(* IEC 61131-3 sources: JingjiangArm/moonboxpro_arm_8.4/Application/Application/任务列表/Main_Task/横向调整处理, 17 files *)

(* ---- StDigitalMicroStepDrive.st ---- *)
(*@CES
Name=StDigitalMicroStepDrive
Type=Gvl
TypeGuid=2db5746d-d284-4425-9f7f-2663a34b0ebc
Guid=10e217d5-ea4e-41f0-93bf-b76d90085cfe
HasDeclaration=True
HasImplementation=False
*)
{DECLARATION}
TYPE StDigitalMicroStepDrive :(*步进电机结构体*)
STRUCT
	xStepDriveEn:BOOL;(*步进电机使能*)
	xStepDriveDir:BOOL;(*步进电机方向*)
	xStepDriveMode:BOOL;(*电机速度位置模式*)(*TRUE 为位置模式，false为速度模式*)
	xStepDriveSpeedMode_Run:BOOL;(*步进电机速度模式启动标志*)
	xStepDriveWorking:BOOL;(*脉冲输出中*)
	xStepDriveAlarm:BOOL;(*步进电机报警*)
	iStepDriveState:INT;(*步进电机状态机*)

	udiStepDriveWorkingTime:UDINT;(*步进电机执行时间*)
	iStepDrivePulsePRev:INT;(*步进电机每圈的脉冲数*)
	iStepDriveNum:INT;(*步进电机减速比分子*)
	iStepDriveDen:INT;(*步进电机减速比分母*)
	lrStepDrivePosPPulse:LREAL;(*步进电机每个脉冲对应的位置值，单位mm*)(*通过测量得到，或者通过计算得到*)
	iStepDriveAccTime_ms:INT;(*步进电机加速时间ms*)
	wStepDrivePulseFre_Sa:WORD;(*步进电机启动脉冲频率*)
	wStepDrivePulseFre_Tar:WORD;(*步进电机目标脉冲频率*)
	wStepDriveAcc_SaToTar:WORD;(*到达目标速度的加速度*)
	wStepDrivePulse:WORD;(*步进电机脉冲数*)
	diStepDrivePluse_Act:DINT;(*步进电机实际走的脉冲数*)
	wStepDrivePulse_Act_Rd_Bak:WORD;(*读取到的步进电机上个周期实际走的脉冲数*)

(*读取模块中的数据*)
	awSpace:ARRAY [1..3] OF WORD;(*W0,W1,W2*)
	wStepDrivePulse_Act_Rd:WORD;(*读取到的步进电机实际走的脉冲数*)(*W3*)
	wStepDriveModuleIOData_Rd:WORD;(*步进电机模块的io输入值*)(*W4*)
	wStepDriveCTL_Rd:WORD;(*读取到的模块的数据*)(*W5*)
(*写入到模块中的参数。规定使用数字量模块 但是plc配置的时候需要配置模拟量模块*)
	wStepDrivePulseFre_Sa_Wr:WORD;(*步进电机启动脉冲频率写入值*)(*W0*)
	wStepDrivePulseFre_Tar_Wr:WORD;(*步进电机目标脉冲频率写入值*)(*W1*)
	wStepDriveAcc_SaToTar_Wr:WORD;(*到达目标速度的加速度写入值*)(*W2*)
	wStepDrivePulse_Wr:WORD;(*步进电机脉冲数写入值*)(*W3*)
	wStepDriveModuleIOData_Wr:WORD;(*步进电机模块的io输出写入*)(*W4*)
	wStepDriveCTL:WORD;(*步进电机控制位*)(*bit9:反馈脉冲数清零(*W5*)
								bit10:脉冲输出标志，1：输出中
								bit11:电机方向
								bit12:速度模式时，高电平输出脉冲，低电平停止输出
								bit13:位置模式时，上升沿开始输出脉冲，脉冲个数到达时停止输出
								bit14:速度、位置模式 0：速度模式，1：位置模式
								bit15:模块使能 0：脉冲输出无效，1：有效
							        *)
END_STRUCT
END_TYPE

{IMPLEMENTATION}

(* ---- StEnc0410R.st ---- *)
(*@CES
Name=StEnc0410R
Type=Gvl
TypeGuid=2db5746d-d284-4425-9f7f-2663a34b0ebc
Guid=6f80462c-d6b3-455f-883a-2142632bafb1
HasDeclaration=True
HasImplementation=False
*)
{DECLARATION}
TYPE StEnc0410R :
STRUCT
	wInputModeCfg:WORD;(*模块输入配置*)
	wInputEncValue:WORD;(*模块输入的编码器个数*)
	wInputEncValue_Bak:WORD;(*上个周期模块输入的编码器个数*)
	diInputEncValue_Total:DINT;(*总的编码器输入个数*)
	diEncValue_Middle:DINT;(*中位临时值*)

	byEnc0410RInPutMode:BYTE;(*模块输入方式选择 0:正交脉冲 1:脉冲+方向 2:正负脉冲*)
	xEnc0410RInPutPulDir:BOOL;(*模块输入脉冲方向 TRUE 取反*)
	byEnc0410RInPutPulCntWay:BYTE;(*模块输入脉冲计数方式 0:z信号开始 1:一直计数*)
	byEncO410RInputVol:BYTE;(*模块输入的电压类型*)

	byEnc0410ROutPutMode:BYTE;(*模块是输出方式选择0:正交脉冲 1:脉冲+方向 2:正负脉冲*)
END_STRUCT
END_TYPE

{IMPLEMENTATION}

(* ---- StStepDriveIOModule.st ---- *)
(*@CES
Name=StStepDriveIOModule
Type=Gvl
TypeGuid=2db5746d-d284-4425-9f7f-2663a34b0ebc
Guid=050a5971-e7ba-4c31-b40e-01a320b97a7e
HasDeclaration=True
HasImplementation=False
*)
{DECLARATION}
TYPE StStepDriveIOModule :
STRUCT
	wIX:WORD;(*输入数据*)(*0：15位为数字量输入*)
	wQX:WORD;(*输出数据*)(*2：9位为数字量继电器输出位*)
END_STRUCT
END_TYPE

{IMPLEMENTATION}

(* ---- TypeEnumEncModule.st ---- *)
(*@CES
Name=TypeEnumEncModule
Type=Gvl
TypeGuid=2db5746d-d284-4425-9f7f-2663a34b0ebc
Guid=5080d035-0ec5-4151-a1b0-b148bbf57879
HasDeclaration=True
HasImplementation=False
*)
{DECLARATION}
TYPE TypeEnumEncModule :
(
	(*0:继电器数字量模块HCB5-1610-DRA*)
	ENCMODULE_HCB5_1610_DRA:=0,
	(*1:Enc0410R模块输出*)
	ENCMODULE_ENC0410R:=1
);
END_TYPE

{IMPLEMENTATION}

(* ---- TypeEnumStepDriveStat.st ---- *)
(*@CES
Name=TypeEnumStepDriveStat
Type=Gvl
TypeGuid=2db5746d-d284-4425-9f7f-2663a34b0ebc
Guid=3c3a1540-5152-4e9f-b7fc-bae736162d3c
HasDeclaration=True
HasImplementation=False
*)
{DECLARATION}
TYPE TypeEnumStepDriveStat :
(
	STEPDRIVE_IDLE,(*空闲*)
	STEPDRIVE_RUN,(*启动*)
	STEPDRIVE_CLR,(*状态清除*)
	STEPDRIVE_WAITING,(*等待一个周期*)
	STEPDRIVE_MODULE_VALID,(*模块使能*)
	STEPDRIVE_PULSEOUT,(*脉冲输出*)
	STEPDRIVE_ALARM(*报警*)
);
END_TYPE

{IMPLEMENTATION}

(* ---- KS_GetEncPluse.st ---- *)
(*@CES
Name=KS_GetEncPluse
Type=FunctionBlock
TypeGuid=6f9dac99-8de1-4efc-8465-68ac443b7d08
Guid=2bf59e22-f994-4ac5-8b2b-a54b74aea4c6
HasDeclaration=True
HasImplementation=True
*)
{DECLARATION}
FUNCTION KS_GetEncPluse : BOOL
VAR_INPUT
	i_pastStDigitalMicroStepDrive :POINTER TO ARRAY [1..MAX_UNIT_NUM] OF StDigitalMicroStepDrive;
	i_pastStEnc0410R:POINTER TO ARRAY [1..MAX_UNIT_NUM] OF StEnc0410R;
END_VAR
VAR
	iN: INT;
END_VAR

{IMPLEMENTATION}
IF i_pastStDigitalMicroStepDrive<>0 AND i_pastStEnc0410R<>0 THEN
	FOR iN:=1 TO MAX_UNIT_NUM BY 1 DO(*针对所有轴进行读取*)
		i_pastStEnc0410R^[iN].wInputEncValue:=
		i_pastStDigitalMicroStepDrive^[iN].wStepDriveModuleIOData_Rd;(*读取回来的编码器脉冲个数，和数字量模块输入公用地址*)

		KS_GetPulse_Act(ADR(i_pastStEnc0410R^[iN].wInputEncValue),
						ADR(i_pastStEnc0410R^[iN].wInputEncValue_Bak),
						ADR(i_pastStEnc0410R^[iN].diInputEncValue_Total) );
	END_FOR
END_IF

(* ---- KS_GetHorizonManuAdj.st ---- *)
(*@CES
Name=KS_GetHorizonManuAdj
Type=FunctionBlock
TypeGuid=6f9dac99-8de1-4efc-8465-68ac443b7d08
Guid=d3a21ffb-1d17-434b-a6db-735f209d6991
HasDeclaration=True
HasImplementation=True
*)
{DECLARATION}
FUNCTION KS_GetHorizonManuAdj : INT(*界面手动调整量2018.9.4.093836*)(*um*)(*返回值为实际需要调整的量，-22222为参数异常*)
(*2022.2.18.164444 按钮方向方向和运动方向相关了*)
(*增加了注释文字@正值是向操作侧@负值是向传动侧@已经和电机旋转方向相关了*)
(*2023.3.9.225628 通过查看动态库发现,动态库中将原来的左按钮赋值为otostudio约定的右按钮
右按钮赋值为otostudio的左按钮
@以前约定向左pabyHorManuBtn= 1 2 5
@向右pabyHorManuBtn=3 4 6
为了不修改动态库,在这里再进行一次取反以保证一致！！@将i_xHorManuDirSwitch=true*)
(*2024.11.6.093600 同步*)
(*2024.11.5.110659*)
(*重新处理界面手动按钮清理，防止整体清除界面手动按钮时B系被A系清理掉了*)
VAR_INPUT
	i_xHorManuDirSwitch:BOOL;(*方向取反*)
	i_iHorManuAdj_Step:INT;(*横向手动调整当量um*)
	i_iHorManuAdj_FastStep:INT;(*横向手动快速调整当量um*)
	i_iHorManuAdj_MidStep:INT;(*横向手动快速调整当量um*)
	piUnitId:POINTER TO INT;(*色组号*)

	pabyHorManuBtn:POINTER TO ARRAY [1..MAX_UNIT_NUM] OF BYTE;(*横向手动按钮，0为不调整，1为左向慢调0.05mm，2为左向快调暂定为0.5mm；3为右向慢调，4为右向快调；
										这里界面上的按钮只控制左右，逻辑控制横向电机是向传动侧还是操作侧运动*)
	padiHorAdjustMent:POINTER TO ARRAY [1..MAX_UNIT_NUM] OF DINT;(*横向手动调整的量*)
	i_iGrpAxisNum_Pu:INT;
	i_abyGrpAxisList: ARRAY [1..MAX_UNIT_NUM] OF BYTE; (*系的轴列表*)
	i_pstStSysParam: POINTER TO StSysParam;
END_VAR
VAR
	iN: INT;
	iCoeff: INT;(*方向系数*)
	iResult: INT;
	iUnitId: INT;
END_VAR

{IMPLEMENTATION}
KS_GetHorizonManuAdj:=0;
IF pabyHorManuBtn<>0 AND padiHorAdjustMent<>0 AND piUnitId<>0 THEN(*指针合法性检查*);
ELSE
	KS_GetHorizonManuAdj:=-22222;(*特殊值标识报警*)
	RETURN;
END_IF

piUnitId^:=0;
IF i_iHorManuAdj_Step<=0 THEN
	i_iHorManuAdj_Step:=50;(*0.05MM*)
ELSE;
END_IF

IF i_iHorManuAdj_FastStep<=0 THEN
	i_iHorManuAdj_FastStep:=500;(*0.5MM*)
ELSE;
END_IF
(*2022.8.9.094516处理0.02档位*)
IF i_iHorManuAdj_MidStep<=0 THEN
	i_iHorManuAdj_FastStep:=100;(*0.1MM*)
ELSE;
END_IF
(*一个周期只处理一个轴*)(*调整量的正值代表向操作侧运动*)
(*2021.10.26.091200  使用轴列表变量*)
FOR iUnitId:=1 TO i_iGrpAxisNum_Pu BY 1 DO(*检查所有色组*)
	iN:=i_abyGrpAxisList[iUnitId];
(*方向*)
	iCoeff:=0;
(*增加0.02档位2022.8.9.094247||*)
(*	IF  pabyHorManuBtn^[iN]=1 OR  pabyHorManuBtn^[iN]=2  THEN(*向左*)*)
	IF  pabyHorManuBtn^[iN]=1 OR  pabyHorManuBtn^[iN]=2 OR  pabyHorManuBtn^[iN]=5 THEN(*向左*)
		IF i_pstStSysParam^.astStUnitParam_UnSave[iN].xMotRev_PrnRoller THEN (*电机反转*)(*向左是向传动侧运动*)
			iCoeff:=-1;
		ELSE(*电机正转*)(*向左是向操作侧运动*)
			iCoeff:=1;
		END_IF
	ELSIF  pabyHorManuBtn^[iN]=3 OR  pabyHorManuBtn^[iN]=4 OR  pabyHorManuBtn^[iN]=6 THEN (*向右*)(*和向左取反*)
		IF i_pstStSysParam^.astStUnitParam_UnSave[iN].xMotRev_PrnRoller THEN (*电机反转*)
			iCoeff:=1;
		ELSE(*电机正转*)
			iCoeff:=-1;
		END_IF
	END_IF

	IF i_xHorManuDirSwitch THEN
		iCoeff:=-iCoeff;
	END_IF
(*调整量值*)
	iResult:=0;
	IF  pabyHorManuBtn^[iN]=1 OR  pabyHorManuBtn^[iN]=3 THEN (*都是慢调*)
		iResult:=(i_iHorManuAdj_Step);
	ELSIF pabyHorManuBtn^[iN]=2 OR  pabyHorManuBtn^[iN]=4 THEN (*都是快调*)
		iResult:=(i_iHorManuAdj_FastStep);
	ELSIF pabyHorManuBtn^[iN]=5 OR  pabyHorManuBtn^[iN]=6 THEN (*中间档位-202022.8.9.094640*)
		iResult:=(i_iHorManuAdj_MidStep);
	END_IF
	iResult:=iResult*iCoeff;

	IF i_pstStSysParam^.astStUnitParam_Save[iN].xLinkage THEN (*检查联动轴*)
		IF pabyHorManuBtn^[iN]<>0 THEN (*说明有调整按下了*)
			pabyHorManuBtn^[iN]:=0;(*清零按钮标志*)(*2024.11.5.110459*)
			KS_GetHorizonManuAdj:=iResult;(*将调整量输出*)
			piUnitId^:=iN;
			padiHorAdjustMent^[iN]:=padiHorAdjustMent^[iN]+iResult;(*在界面显示*)
			EXIT;
		END_IF
	ELSE
		pabyHorManuBtn^[iN]:=0;(*清零按钮标志*)(*2024.11.5.110459*)
	END_IF
END_FOR

(* ---- KS_GetPulse_Act.st ---- *)
(*@CES
Name=KS_GetPulse_Act
Type=FunctionBlock
TypeGuid=6f9dac99-8de1-4efc-8465-68ac443b7d08
Guid=7e51e991-78cc-4457-be42-c8156f7134b7
HasDeclaration=True
HasImplementation=True
*)
{DECLARATION}
FUNCTION KS_GetPulse_Act : int
VAR_INPUT
	pwStepDrivePulse_Act_Rd :POINTER TO WORD;(*读取到的脉冲数*)
	pwStepDrivePulse_Act_Rd_Bak:POINTER TO WORD;(*上个周期读到的脉冲数*)
	pdiStepDrivePulse_Act:POINTER TO DINT;(*实际走的脉冲数*)
END_VAR
VAR
	iStepDrivePulse_Act_Rd: INT;
	iStepDrivePulse_Act_Rd_Bak: INT;
	iDeltaPulse: INT;(*步进电机脉冲变化量*)
END_VAR

{IMPLEMENTATION}
KS_GetPulse_Act:=0;
IF pwStepDrivePulse_Act_Rd<>0 AND pwStepDrivePulse_Act_Rd_Bak<>0 AND pdiStepDrivePulse_Act <>0 THEN;
ELSE
	KS_GetPulse_Act:=-1;
	RETURN;
END_IF

iStepDrivePulse_Act_Rd:=WORD_TO_INT(pwStepDrivePulse_Act_Rd^);
iStepDrivePulse_Act_Rd_Bak:= WORD_TO_INT(pwStepDrivePulse_Act_Rd_Bak^);

IF iStepDrivePulse_Act_Rd <> iStepDrivePulse_Act_Rd_Bak THEN
	iDeltaPulse:=(iStepDrivePulse_Act_Rd-iStepDrivePulse_Act_Rd_Bak);
	pdiStepDrivePulse_Act^:=pdiStepDrivePulse_Act^+iDeltaPulse;
ELSE;
END_IF

pwStepDrivePulse_Act_Rd_Bak^:=INT_TO_WORD(iStepDrivePulse_Act_Rd);(*保存上个周期的值*)

(* ---- KS_SetStepDriveModulePara.st ---- *)
(*@CES
Name=KS_SetStepDriveModulePara
Type=FunctionBlock
TypeGuid=6f9dac99-8de1-4efc-8465-68ac443b7d08
Guid=21a3679d-2e4f-4802-b9d7-d00f676e215d
HasDeclaration=True
HasImplementation=True
*)
{DECLARATION}
FUNCTION KS_SetStepDriveModulePara : BOOL(*设置步进电机脉冲输出模块脉冲方式参数*)
(*2019.5.15.112350|liu.yt|必须放在KS_FB_StepDriveCTL后执行，KS_FB_StepDriveCTL会清零，功能块再次再次赋值，反之则无效赋值*)
(*2019.4.18.130455 增加了ENCO410R型模块输入输出控制参数,主要用于高速编码器输入输出控制。MHZ频率*)
VAR_INPUT
	i_xMultiple_Input: BOOL;(*参数输入方式选择：多参数 或者 单参数*)
	i_byEncO410RInputVol:BYTE;(*模块输入的电压类型选择：0 是5v；1是24v*)
	i_byEnc0410RInPutMode:BYTE;(*模块输入方式选择 0:正交脉冲 1:脉冲+方向 2:正负脉冲*)
	i_xEnc0410RInPutPulDir:BOOL;(*模块输入脉冲方向 TRUE 取反*)
	i_byEnc0410RInPutPulCntWay:BYTE;(*模块输入脉冲计数方式 0:z信号开始 1:一直计数*)

	i_byEnc0410ROutPutMode:BYTE;(*模块输出方式选择 0:正交脉冲 1:脉冲+方向 2:正负脉冲*)
	i_pastStDigitalMicroStepDrive :POINTER TO ARRAY [1..MAX_UNIT_NUM] OF StDigitalMicroStepDrive;
	i_pastStEnc0410R:POINTER TO ARRAY [1..MAX_UNIT_NUM] OF StEnc0410R;
END_VAR
VAR
(*bit7:8 脉冲输出模式，仅限于EncO410R模块，0:正交脉冲 1:脉冲+方向 2:正负脉冲*)
	wEncO410ROutPutMode_ClrCtlBit:WORD:=16#FE7F;(*利用与运算清除7:8位*)
(*利用或运算定义控制位*)
	wEncO410ROutPutMode_QuadPul:WORD:=0;		(*正交脉冲输出模式	bit 7:8=0*)
	wEncO410ROutPutMode_PulAndDir:WORD:=16#0080;	(*脉冲+方向输出模式	bit 7:8=1*)
	wEncO410ROutPutMode_PlusMinusPul:WORD:=16#0100;(*正负脉冲输出模式	bit 7:8=2*)

(*************************************************)
(*Enc0410R 模块输入配置*)(*bit0:1 脉冲输入模式。bit2 方向取反。bit3 计数模式*)
	wEncO410RInPutMode_ClrCtlBit:WORD:=16#FFF0;(*利用与运算清除低四位*)
(*利用或运算定义控制位*)
	wEncO410RInPutMode_QuadPul:WORD:=0;		(*正交脉冲输出模式	bit 0:1=0*)
	wEncO410RInPutMode_PulAndDir:WORD:=16#0001;	(*脉冲+方向输出模式	bit 0:1=1*)
	wEncO410RInPutMode_PlusMinusPul:WORD:=16#0002;(*正负脉冲输出模式	bit 0:1=2*)
	wEncO410RInPutMode_PlusDir:WORD:=16#0004;(*bit2 脉冲方向*)
(*	wEncO410RInPutMode_PlusCntWay_Z:WORD:=0;(*脉冲计数模式：z信号开始*)*)
	wEncO410RInPutMode_PlusCntWay_All:WORD:=16#0008;(*脉冲计数模式：一直计数*)
	wEncO410RInPutMode_Vol:WORD:=16#0010;(*bit4 电压输入类型 0 是5v；1是24v*)

	iN: INT;
	wStepDriveCTL: WORD;
	wEncO410RInPutModeCfg: WORD;

	byEnc0410RInPutMode:BYTE;(*模块输入方式选择 0:正交脉冲 1:脉冲+方向 2:正负脉冲*)
	xEnc0410RInPutPulDir:BOOL;(*模块输入脉冲方向 TRUE 取反*)
	byEnc0410RInPutPulCntWay:BYTE;(*模块输入脉冲计数方式 0:z信号开始 1:一直计数*)
	byEncO410RInputVol: BYTE;(*模块输入的电压类型选择：0 是5v；1是24v*)

	byEnc0410ROutPutMode:BYTE;(*模块输出方式选择 0:正交脉冲 1:脉冲+方向 2:正负脉冲*)
END_VAR

{IMPLEMENTATION}
IF i_pastStDigitalMicroStepDrive<>0 AND i_pastStEnc0410R<>0 THEN
	FOR iN:=1 TO MAX_UNIT_NUM BY 1 DO(*针对所有轴进行控制*)
		IF i_xMultiple_Input THEN(*多参数输入*)
			byEnc0410RInPutMode:=i_pastStEnc0410R^[iN].byEnc0410RInPutMode;
			xEnc0410RInPutPulDir:=i_pastStEnc0410R^[iN].xEnc0410RInPutPulDir;
			byEnc0410RInPutPulCntWay:=i_pastStEnc0410R^[iN].byEnc0410RInPutPulCntWay;
			byEncO410RInputVol:=i_pastStEnc0410R^[iN].byEncO410RInputVol;
			byEnc0410ROutPutMode:=i_pastStEnc0410R^[iN].byEnc0410ROutPutMode;
		ELSE(*单参数输入*)
			byEnc0410RInPutMode:=i_byEnc0410RInPutMode;
			xEnc0410RInPutPulDir:=i_xEnc0410RInPutPulDir;
			byEnc0410RInPutPulCntWay:=i_byEnc0410RInPutPulCntWay;
			byEncO410RInputVol:=i_byEncO410RInputVol;
			byEnc0410ROutPutMode:=i_byEnc0410ROutPutMode;
		END_IF

		(*脉冲输出配置*)
		wStepDriveCTL:=i_pastStDigitalMicroStepDrive^[iN].wStepDriveCTL;
		wStepDriveCTL:=wStepDriveCTL AND wEncO410ROutPutMode_ClrCtlBit;(*清零相应位*)
		(*输出方式配置*)
		CASE byEnc0410ROutPutMode OF
		1:(*脉冲+方向*)
			wStepDriveCTL:=wStepDriveCTL+wEncO410ROutPutMode_PulAndDir;
		2:(*正负脉冲*)
			wStepDriveCTL:=wStepDriveCTL+wEncO410ROutPutMode_PlusMinusPul;
		ELSE(*默认输出方式是正交脉冲*)
			wStepDriveCTL:=wStepDriveCTL+wEncO410ROutPutMode_QuadPul;
		END_CASE

		i_pastStDigitalMicroStepDrive^[iN].wStepDriveCTL:=wStepDriveCTL;

		(*脉冲输入配置*)
		(*Enc0410R的输入参数配置和继电器数字量模块公用IO输入输出地址*)
		wEncO410RInPutModeCfg:=0;

		(*输入方式配置*)

		CASE byEnc0410RInPutMode OF
		1:(*脉冲+方向*)
			wEncO410RInPutModeCfg:=wEncO410RInPutModeCfg+wEncO410RInPutMode_PulAndDir;
		2:(*正负脉冲*)
			wEncO410RInPutModeCfg:=wEncO410RInPutModeCfg+wEncO410RInPutMode_PlusMinusPul;
		ELSE(*默认输出方式是正交脉冲*)
			wEncO410RInPutModeCfg:=wEncO410RInPutModeCfg+wEncO410RInPutMode_QuadPul;
		END_CASE

		(*方向取反*)
		IF xEnc0410RInPutPulDir THEN wEncO410RInPutModeCfg:=wEncO410RInPutModeCfg+wEncO410RInPutMode_PlusDir;END_IF

		(*计数方式选择*)
		IF byEnc0410RInPutPulCntWay<>0 THEN wEncO410RInPutModeCfg:=wEncO410RInPutModeCfg+wEncO410RInPutMode_PlusCntWay_All;END_IF

		(*输入电压类型 0 是5v  1是24v*)
		IF byEncO410RInputVol=1 THEN wEncO410RInPutModeCfg:=wEncO410RInPutModeCfg+wEncO410RInPutMode_Vol;END_IF

		i_pastStEnc0410R^[iN].wInputModeCfg:=wEncO410RInPutModeCfg;
	END_FOR
END_IF

(* ---- KS_FB_AxisHorAdj.st ---- *)
(*@CES
Name=KS_FB_AxisHorAdj
Type=FunctionBlock
TypeGuid=6f9dac99-8de1-4efc-8465-68ac443b7d08
Guid=bd4bc8d3-26df-4dfe-bfb9-1ac44a7e80cd
HasDeclaration=True
HasImplementation=True
*)
{DECLARATION}
FUNCTION_BLOCK KS_FB_AxisHorAdj(*从站横向*)
(*2022.6.10.161033 修复横向运动限位问题*)
(*屏蔽使用移动到KS_FB_GrpHorAdj函数中*)
(*2025.4.20.104124从站横向运动功能，停机状态取消联动相关|开机状态下非联动轴也可以运动*)
(*已经不使用了@@@@*)
VAR_INPUT
	i_xEn									: BOOL;(*功能块使能*)
	i_iGrpAxisNum_Pu						: INT; (*色组轴数*)
	i_aiGrpAxisList							: ARRAY [1..MAX_UNIT_NUM] OF INT; (*系的轴列表*)
	i_pastStIOMap_AxisBasic					: POINTER TO ARRAY [1..MAX_UNIT_NUM] OF StIOMap_Axis_FE; (*基础io|*)
	i_xFlag_Estop							: BOOL;(*急停标志*)
	i_xFlag_Stop							: BOOL;(*停机标志*)
	i_lrVel_HorzPreRegister					: LREAL;
	i_lrVel_HorzAdjust						: LREAL;
	i_iCycleTime_Plc						: INT;
	i_pastStAxisRapidAdjProf_H				: POINTER TO ARRAY [1..MAX_UNIT_NUM] OF StAxisRapidAdjProf_H;(*纵向快速对版|*)
	i_pstStSysParam: POINTER TO StSysParam;
	i_iGrpId: INT;
END_VAR
VAR_OUTPUT

	o_axAxisHorAdjing: ARRAY [1..MAX_UNIT_NUM] OF BOOL;
END_VAR
VAR
	iN: INT;
	iUnitId: INT;
	//pstStAxisParam: POINTER TO StAxisParam;
	pstStIOMap_AxisBasic: POINTER TO StIOMap_Axis_FE;

	lrAdjustVal_H_PerCycle: LREAL;
	axAxisHorAdjSts: ARRAY [1..MAX_UNIT_NUM] OF BOOL;
	axAxisHorAdj_End: ARRAY [1..MAX_UNIT_NUM] OF BOOL;
	iRtn: INT;
	iAdjustment_HorAxisAdj: INT;
	axHorAxisAdjStop: ARRAY [1..MAX_UNIT_NUM] OF BOOL;
	axHorAxisAdjStart: ARRAY [1..MAX_UNIT_NUM] OF BOOL;
	xFlag_HorAxisAdj: BOOL;
	wSts_HorzManuPreReg:WORD;
	xAutoMove_H: BOOL;(*2025.4.20.110020+*)
END_VAR

{IMPLEMENTATION}
IF i_xEn AND
	(i_iGrpAxisNum_Pu>=1 AND i_iGrpAxisNum_Pu<=MAX_UNIT_NUM) AND
	i_pastStIOMap_AxisBasic<>0 AND
	i_pastStAxisRapidAdjProf_H<>0 THEN(*2019.11.18.153726_*)

	FOR iN:= 1 TO i_iGrpAxisNum_Pu BY 1 DO
		iUnitId:= i_aiGrpAxisList[iN];
		pstStIOMap_AxisBasic:= ADR(i_pastStIOMap_AxisBasic^[iUnitId]);

		(*--------------------------------------------------|2019.11.18.153930_*)
		(*横向快速对版改成单个轴处理时放在循环内处理|*)
		iRtn:= KS_FetchRapidAdjValue_H(i_pastStAxisRapidAdjProf_H, iUnitId, ADR(iAdjustment_HorAxisAdj));
		(*2025.4.20.110359 同步*)
		(*2024.01.17.161205 增加清除处理*)
		axHorAxisAdjStart[iUnitId]:= FALSE;
		axHorAxisAdjStop[iUnitId]:= FALSE;
		IF iRtn=0 THEN
			IF iAdjustment_HorAxisAdj=-32767 THEN(*人为停止标志|*)
				axHorAxisAdjStop[iUnitId]:= TRUE;
				axHorAxisAdjStart[iUnitId]:= FALSE;
			ELSIF iAdjustment_HorAxisAdj<>0 THEN
				axHorAxisAdjStop[iUnitId]:= FALSE;
				axHorAxisAdjStart[iUnitId]:= TRUE;
				i_pstStSysParam^.astStUnitParam_UnSave[iUnitId].alrTotalAdjustVal_ManuCoarse_vh[2]:= i_pstStSysParam^.astStUnitParam_UnSave[iUnitId].alrTotalAdjustVal_ManuCoarse_vh[2]+iAdjustment_HorAxisAdj;
			END_IF
		END_IF

		IF (NOT i_xFlag_Estop) (*AND i_xFlag_Stop*) THEN(*非急停*)
			(*2025.4.20.105720 修改条件*)
			IF i_xFlag_Stop THEN(*不用限制单联动*)
				xAutoMove_H:=TRUE;
			ELSE(*非停机状态下|只有单动的可以*)
				xAutoMove_H:=NOT i_pstStSysParam^.astStUnitParam_Save[iUnitId].xLinkage;
			END_IF

			IF (*pstStAxisParam^.xLinkage*)xAutoMove_H THEN
				IF axHorAxisAdjStart[iUnitId] AND (NOT axAxisHorAdjSts[iUnitId]) THEN(*开始运行*)
					axAxisHorAdjSts[iUnitId]:= TRUE;
					axHorAxisAdjStart[iUnitId]:= FALSE;
				END_IF
				IF axHorAxisAdjStop[iUnitId] AND axAxisHorAdjSts[iUnitId] THEN(*停止运行*)
					axAxisHorAdjSts[iUnitId]:= FALSE;
					axHorAxisAdjStop[iUnitId]:= FALSE;
				END_IF
			ELSE
				axHorAxisAdjStart[iUnitId]:= FALSE;
				axHorAxisAdjStop[iUnitId]:= FALSE;
				axAxisHorAdjSts[iUnitId]:= FALSE;
				IF i_pstStSysParam^.astStUnitParam_UnSave[iUnitId].alrTotalAdjustVal_ManuCoarse_vh[2]<>0 THEN
					i_pstStSysParam^.astStUnitParam_UnSave[iUnitId].alrTotalAdjustVal_ManuCoarse_vh[2]:= 0;
				END_IF

			END_IF
		ELSE(*2019.11.20.115512 增加了清除axHorAxisAdjStart
								axHorAxisAdjStop标志|Liu.yt*)
			axHorAxisAdjStart[iUnitId]:= FALSE;
			axHorAxisAdjStop[iUnitId]:= FALSE;
			IF axAxisHorAdjSts[iUnitId] THEN
				axAxisHorAdjSts[iUnitId]:= FALSE;(*急停或者非停机-直接停止运行*)
				i_pstStSysParam^.astStUnitParam_UnSave[iUnitId].alrTotalAdjustVal_ManuCoarse_vh[2]:= 0;
			END_IF
		END_IF

		IF pstStIOMap_AxisBasic^.o_xRel_Press OR (NOT pstStIOMap_AxisBasic^.i_xHorzMotor_FastSpd) THEN
		(*快调/慢调处理*)
			lrAdjustVal_H_PerCycle:= i_lrVel_HorzAdjust*INT_TO_LREAL(i_iCycleTime_Plc);
		ELSE
			lrAdjustVal_H_PerCycle:= i_lrVel_HorzPreRegister*INT_TO_LREAL(i_iCycleTime_Plc);
		END_IF

		IF axAxisHorAdjSts[iUnitId] THEN (*色组进入到横向对版状态*)
			xFlag_HorAxisAdj:= TRUE;

			(*2025.4.20.105821 屏蔽联动条件*)
			IF i_pstStSysParam^.astStUnitParam_Save[iUnitId].xLinkage OR TRUE THEN(*色组联动*)
				IF NOT axAxisHorAdj_End[iUnitId] THEN
					IF NOT o_axAxisHorAdjing[iUnitId] THEN
						o_axAxisHorAdjing[iUnitId]:= TRUE;
						(*横向对版量叠加到横向手动粗调仓库*)
						i_pstStSysParam^.astStUnitParam_UnSave[iUnitId].alrTotalAdjustVal_ManuCoarse_vh[2]:= -i_pstStSysParam^.astStUnitParam_UnSave[iUnitId].alrTotalAdjustVal_ManuCoarse_vh[2]*1000;(*单位um*)
					ELSE
(*2022.6.10.160946*)
(*
						IF pstStIOMap_AxisBasic^.i_xPosLimit_Left OR pstStIOMap_AxisBasic^.i_xPosLimit_Right THEN (*到达左右限位，直接清零调整量*)
							pstStAxisParam^.alrTotalAdjustVal_ManuCoarse_vh[2]:= 0;
						END_IF
*)

						IF (pstStIOMap_AxisBasic^.i_xPosLimit_Right AND i_pstStSysParam^.astStUnitParam_UnSave[iUnitId].alrTotalAdjustVal_ManuCoarse_vh[2]<0) OR
							(pstStIOMap_AxisBasic^.i_xPosLimit_Left AND i_pstStSysParam^.astStUnitParam_UnSave[iUnitId].alrTotalAdjustVal_ManuCoarse_vh[2]>0) THEN
							i_pstStSysParam^.astStUnitParam_UnSave[iUnitId].alrTotalAdjustVal_ManuCoarse_vh[2]:=0;
						END_IF

						IF i_pstStSysParam^.astStUnitParam_UnSave[iUnitId].alrTotalAdjustVal_ManuCoarse_vh[2]=0 THEN(*调整量消耗完成*)
							o_axAxisHorAdjing[iUnitId]:= FALSE;
							axAxisHorAdj_End[iUnitId]:= TRUE;
							axAxisHorAdjSts[iUnitId]:= FALSE;
						END_IF
					END_IF
				END_IF
			ELSE(*单动*)
				o_axAxisHorAdjing[iUnitId]:= FALSE;
				axAxisHorAdj_End[iUnitId]:= TRUE;
				axAxisHorAdjSts[iUnitId]:= FALSE;
				IF i_pstStSysParam^.astStUnitParam_UnSave[iUnitId].alrTotalAdjustVal_ManuCoarse_vh[2]<>0 THEN
					i_pstStSysParam^.astStUnitParam_UnSave[iUnitId].alrTotalAdjustVal_ManuCoarse_vh[2]:=0;
				END_IF
			END_IF
		ELSE
			IF xFlag_HorAxisAdj THEN
				xFlag_HorAxisAdj:= FALSE;
			END_IF
			o_axAxisHorAdjing[iUnitId]:= FALSE;
			axAxisHorAdj_End[iUnitId]:= FALSE;
			IF i_pstStSysParam^.astStUnitParam_UnSave[iUnitId].alrTotalAdjustVal_ManuCoarse_vh[2]<>0 THEN(*退出横向对版状态，调整量清零*)
				i_pstStSysParam^.astStUnitParam_UnSave[iUnitId].alrTotalAdjustVal_ManuCoarse_vh[2]:=0;
			END_IF
		END_IF

		IF axAxisHorAdjSts[iUnitId] THEN
			IF ABS(i_pstStSysParam^.astStUnitParam_UnSave[iUnitId].alrTotalAdjustVal_ManuCoarse_vh[2])>lrAdjustVal_H_PerCycle THEN
				IF i_pstStSysParam^.astStUnitParam_UnSave[iUnitId].alrTotalAdjustVal_ManuCoarse_vh[2]>0 THEN
					(*正向*)
					i_pstStSysParam^.astStUnitParam_UnSave[iUnitId].alrCurCycleAdjustVal_ManuCoarse_vh[2]:= lrAdjustVal_H_PerCycle;
					i_pstStSysParam^.astStUnitParam_UnSave[iUnitId].alrTotalAdjustVal_ManuCoarse_vh[2]:= i_pstStSysParam^.astStUnitParam_UnSave[iUnitId].alrTotalAdjustVal_ManuCoarse_vh[2] - i_pstStSysParam^.astStUnitParam_UnSave[iUnitId].alrCurCycleAdjustVal_ManuCoarse_vh[2];
					i_pstStSysParam^.astStUnitParam_UnSave[iUnitId].axCurCycleAdjustVal_ManuCoarse_done_vh[2]:= FALSE;
					pstStIOMap_AxisBasic^.o_xHorzMotor_CW:= TRUE;(*正转*)
					pstStIOMap_AxisBasic^.o_xHorzMotor_CCW:= FALSE;
				ELSE
					(*反向*)
					i_pstStSysParam^.astStUnitParam_UnSave[iUnitId].alrCurCycleAdjustVal_ManuCoarse_vh[2]:= -lrAdjustVal_H_PerCycle;
					i_pstStSysParam^.astStUnitParam_UnSave[iUnitId].alrTotalAdjustVal_ManuCoarse_vh[2]:= i_pstStSysParam^.astStUnitParam_UnSave[iUnitId].alrTotalAdjustVal_ManuCoarse_vh[2] - i_pstStSysParam^.astStUnitParam_UnSave[iUnitId].alrCurCycleAdjustVal_ManuCoarse_vh[2];
					i_pstStSysParam^.astStUnitParam_UnSave[iUnitId].axCurCycleAdjustVal_ManuCoarse_done_vh[2]:= FALSE;
					pstStIOMap_AxisBasic^.o_xHorzMotor_CCW:= TRUE;(*反转*)
					pstStIOMap_AxisBasic^.o_xHorzMotor_CW:= FALSE;
				END_IF
			ELSE
				IF o_axAxisHorAdjing[iUnitId] THEN
					i_pstStSysParam^.astStUnitParam_UnSave[iUnitId].alrTotalAdjustVal_ManuCoarse_vh[2]:= 0;
				END_IF
				pstStIOMap_AxisBasic^.o_xHorzMotor_CW:= FALSE;
				pstStIOMap_AxisBasic^.o_xHorzMotor_CCW:= FALSE;
			END_IF

		END_IF
(*往从站发送*)
		i_pstStSysParam^.astStUnitParam_UnSave[iUnitId].iPos_HorzManuPreReg:= -LREAL_TO_INT(i_pstStSysParam^.astStUnitParam_UnSave[iUnitId].alrTotalAdjustVal_ManuCoarse_vh[2]/1000);

		wSts_HorzManuPreReg.0:= o_axAxisHorAdjing[iUnitId];
		wSts_HorzManuPreReg.1:= pstStIOMap_AxisBasic^.o_xHorzMotor_CW;
		wSts_HorzManuPreReg.2:= pstStIOMap_AxisBasic^.o_xHorzMotor_CCW;
		wSts_HorzManuPreReg.3:= pstStIOMap_AxisBasic^.i_xPosLimit_Left;
		wSts_HorzManuPreReg.4:= pstStIOMap_AxisBasic^.i_xPosLimit_Right;
		wSts_HorzManuPreReg.5:= i_pstStSysParam^.astStGrpParam_UnSave[i_iGrpId].xFlag_Stop;

		i_pstStSysParam^.astStUnitParam_UnSave[iUnitId].wSts_HorzManuPreReg:= wSts_HorzManuPreReg;
	END_FOR

END_IF

(* ---- KS_FB_Debug_Get_mmPpul.st ---- *)
(*@CES
Name=KS_FB_Debug_Get_mmPpul
Type=FunctionBlock
TypeGuid=6f9dac99-8de1-4efc-8465-68ac443b7d08
Guid=61707722-1ee3-4896-b414-72dee3b67cb6
HasDeclaration=True
HasImplementation=True
*)
{DECLARATION}
FUNCTION_BLOCK KS_FB_Debug_Get_mmPpul(*调试模式下计算出的每个脉冲对应的位置值单位mm/pul*)
VAR_INPUT
	i_xEn:BOOL;(*功能块使能*)
	i_xStartTrig:BOOL;(*启动步进电机*)
	i_xCalEn:BOOL;(*计算使能标志*)
	i_iNum:INT;(*执行该动作的色组号*)
	i_iStepDriveSa_Vel:INT;(*步进电机启动速度*)
	i_iStepDrivePreReg_Vel:INT;(*z步进电机预套速度R/MIN*)
	i_diPulse:DINT;(*执行的脉冲数pul*)
	i_lrPos_Act:LREAL;(*实际走的距离mm*)
	i_pastStDigitalMicroStepDrive :POINTER TO ARRAY [1..MAX_UNIT_NUM] OF StDigitalMicroStepDrive;
END_VAR
VAR_OUTPUT
	o_xEn:BOOL;(**)
	o_xDebugTestDone: BOOL;(*测试完成了*)
	o_lrResult:LREAL;(*计算出的结果*)(*只有效一个周期*)
	o_iErrCode: INT;(*-1 地址错误。-2 数组下标越界,-3 输入参数错误*)
END_VAR
VAR
	xPreStartTrig: BOOL;(*用来控制启动检测按钮的上升沿*)
	stStDigitalMicroStepDrive_Temp: StDigitalMicroStepDrive;
	lrTemp: LREAL;
	lrTemp1: LREAL;
	xDebugTesting: BOOL;(*处于测试状态中*)
	xPreStepDriveWorking: BOOL;(*用来检测脉冲输出下降沿*)
	xPreCalEn: BOOL;(*用于检测计算使能上升沿*)
END_VAR

{IMPLEMENTATION}
(*输入参数检查*)
o_iErrCode:=0;
o_lrResult:=0;
IF i_pastStDigitalMicroStepDrive<>0 THEN;
ELSE
	o_iErrCode:=-1;
	RETURN;
END_IF

IF i_iNum>=1 AND i_iNum<=MAX_UNIT_NUM THEN
;
ELSE
	i_iNum:=1;
	o_iErrCode:=-2;
END_IF

IF ABS(i_diPulse)>65535 AND i_diPulse<>0 THEN
	i_diPulse:=65535*i_diPulse/i_diPulse;
	o_iErrCode:=-3;
END_IF

IF i_lrPos_Act<0 THEN
	i_lrPos_Act:=ABS(i_lrPos_Act);
	o_iErrCode:=-3;
END_IF

IF i_iStepDriveSa_Vel<0 THEN
	i_iStepDriveSa_Vel:=ABS(i_iStepDriveSa_Vel);
	o_iErrCode:=-3;
END_IF

IF i_iStepDrivePreReg_Vel<0 THEN
	i_iStepDrivePreReg_Vel:=ABS(i_iStepDrivePreReg_Vel);
	o_iErrCode:=-3;
END_IF

stStDigitalMicroStepDrive_Temp:=i_pastStDigitalMicroStepDrive^[i_iNum];
IF i_xEn THEN(*使能计算*)
	IF i_xStartTrig  AND NOT xPreStartTrig THEN(*检测按钮上升沿*)
		IF NOT xDebugTesting THEN
			o_xDebugTestDone:=FALSE;
			lrTemp:=i_pastStDigitalMicroStepDrive^[i_iNum].iStepDrivePulsePRev*i_iStepDriveSa_Vel/60.0;(*pul/s*)
			lrTemp1:=i_pastStDigitalMicroStepDrive^[i_iNum].iStepDrivePulsePRev*i_iStepDrivePreReg_Vel/60.0;(*pul/s*)
			IF i_pastStDigitalMicroStepDrive^[i_iNum].iStepDriveState=STEPDRIVE_IDLE  THEN(*空闲状态*)
				i_pastStDigitalMicroStepDrive^[i_iNum].iStepDriveState:=STEPDRIVE_RUN;(*启动步进电机调整*)
				i_pastStDigitalMicroStepDrive^[i_iNum].wStepDrivePulseFre_Sa:=LREAL_TO_WORD(lrTemp);
				i_pastStDigitalMicroStepDrive^[i_iNum].wStepDrivePulseFre_Tar:=LREAL_TO_WORD(lrTemp1);
				i_pastStDigitalMicroStepDrive^[i_iNum].wStepDrivePulse:=DINT_TO_WORD(ABS(i_diPulse));(*写入的脉冲数*)
				i_pastStDigitalMicroStepDrive^[i_iNum].xStepDriveMode:=TRUE;(*位置模式*)
				i_pastStDigitalMicroStepDrive^[i_iNum].xStepDriveSpeedMode_Run:=FALSE;(*置位速度模式输出标志*)
				IF i_diPulse>0 THEN
					i_pastStDigitalMicroStepDrive^[i_iNum].xStepDriveDir:=TRUE;(*为正值的时候我们认为是向传动侧转动，由于默认方向是向操作侧转动，故写为true*)
				ELSE
					i_pastStDigitalMicroStepDrive^[i_iNum].xStepDriveDir:=FALSE;(*为负值的时候我们认为是向操作侧转动，由于默认方向是向操作侧转动，故写为false*)
				END_IF
			END_IF
		ELSE(*再次按下启动按钮我们就退出测试位置的状态*);
			i_pastStDigitalMicroStepDrive^[i_iNum].iStepDriveState:=STEPDRIVE_IDLE;(*先退出到空闲状态*)
		END_IF
		xDebugTesting:=NOT xDebugTesting;
	END_IF

	IF xDebugTesting THEN (*已经处于测试的状态了,这个时候需要一直检测是否执行完成了*)
		IF NOT i_pastStDigitalMicroStepDrive^[i_iNum].xStepDriveWorking AND  xPreStepDriveWorking THEN(*脉冲输出标志下降沿*)
			i_pastStDigitalMicroStepDrive^[i_iNum].iStepDriveState:=STEPDRIVE_IDLE;(*退出到空闲状态*)
			xDebugTesting:=FALSE;
			o_xDebugTestDone:=TRUE;
		END_IF
	ELSE;
	END_IF

	IF o_xDebugTestDone THEN (*测试完成 接着我们计算每个脉冲对应的位置值*)
		IF i_xCalEn AND NOT xPreCalEn THEN(*计算上升沿标志*)
			IF i_pastStDigitalMicroStepDrive^[i_iNum].diStepDrivePluse_Act<>0 THEN
				o_lrResult:=ABS(i_lrPos_Act/i_pastStDigitalMicroStepDrive^[i_iNum].diStepDrivePluse_Act);
			ELSE
				o_iErrCode:=-4;
			END_IF
		END_IF
	END_IF
ELSE
	xDebugTesting:=FALSE;
	o_xDebugTestDone:=FALSE;
END_IF
xPreStepDriveWorking:=i_pastStDigitalMicroStepDrive^[i_iNum].xStepDriveWorking;
xPreStartTrig:=i_xStartTrig;
xPreCalEn:=i_xCalEn;

(* ---- KS_FB_GrpHorAdj.st ---- *)
(*@CES
Name=KS_FB_GrpHorAdj
Type=FunctionBlock
TypeGuid=6f9dac99-8de1-4efc-8465-68ac443b7d08
Guid=d546f829-7451-435f-8672-15bc73f9dc0f
HasDeclaration=True
HasImplementation=True
*)
{DECLARATION}
FUNCTION_BLOCK KS_FB_GrpHorAdj(*传统横向电机调整*)
(*2023.3.8.214754
移植KS_FB_AxisHorAdj 代码
程序逻辑只有操作侧和传动侧的方向
@位置正值代表向操作侧运动
@位置负值代表向传动侧运动
电机输出只有正转和反转
@正转是向操作侧
@反转是向传动侧*)
(*2023.3.10.105606 为了兼容外部的硬件限位处理
这里将限位定义调整下
@i_xMove_Left 为正转限位即操作侧限位
@i_xMove_Right 为反转限位即传动侧限位
@支持密码切换将限位定义切换为左右限位@dwControlComplexBits.17|未处理密码切换部分*)

(*2024.01.17.162016 优化从站横向控制标志处理@现场偶尔出现从站横向操作无响应问题*)
(*2025.4.20.104124从站横向运动功能，停机状态取消联动相关|开机状态下非联动轴也可以运动*)
(*2025.9.5.104845 自动横向调整时单周期调整量超过1丝的量不会因为自动速度太快而不响应@现场会出现小误差一直不能回来(单个周期的调整量太大了)*)
VAR_INPUT
	i_xEn: BOOL;(*使能*)
	i_iGrpAxisNum_Pu: INT; (*色组轴数*)
	i_abyGrpAxisList: ARRAY [1..MAX_UNIT_NUM] OF BYTE; (*系的轴列表*)
	i_pastStIOMap_AxisBasic: POINTER TO ARRAY [1..MAX_UNIT_NUM] OF StIOMap_Axis_FE; (*基础io|*)
	i_pastStIOMap_AxisExtra: POINTER TO ARRAY [1..MAX_UNIT_NUM] OF StIOMap_Axis_Extra_FE; (* 扩展io|*)
	i_lrVel_HorzAdjust		: LREAL;(*mm/s; um/ms; 横向调整速度|*)
	i_lrVel_HorzPreRegister		: LREAL;(*mm/s;横向预套准速度|*)
	(*2023.3.8.114628*)
	i_xFlag_Estop							: BOOL;(*急停标志*)
	i_xFlag_Stop							: BOOL;(*停机标志*)
	i_iCycleTime_Plc						: INT;
	i_pastStAxisRapidAdjProf_H				: POINTER TO ARRAY [1..MAX_UNIT_NUM] OF StAxisRapidAdjProf_H;(*纵向快速对版|*)
	i_pstStSysParam: POINTER TO StSysParam;
	i_xHorLimit:BOOL;(*横向限位定义修改为左右|默认是纤维定义为正反方向*)
	i_iGrpId: INT;
	i_xHorManuCtrl:BOOL;(*界面横向手动修正功能*)
END_VAR
VAR_OUTPUT
	o_xEno: BOOL;
	o_iErNo: INT;(*0成功\-1参数失败|*)
	o_axAxisHorAdjing: ARRAY [1..MAX_UNIT_NUM] OF BOOL;
END_VAR
VAR
	iN: INT;

	iUnitId: INT;

	pstStIOMap_AxisBasic: POINTER TO StIOMap_Axis_FE;
	pstStIOMap_AxisExtra: POINTER TO StIOMap_Axis_Extra_FE;
	//pstStAxisParam: POINTER TO StAxisParam;

	xFlag_PreRegister_H: BOOL;(*用来表征是否进入过横向预套准状态*)

	wHorzMotorDir: WORD;(*.0 |正转方向
					.1|反转方向*)
	awPreHorzMotorDir: ARRAY [1..MAX_UNIT_NUM] OF WORD;
	axHorzMotorStart_Delay: ARRAY [1..MAX_UNIT_NUM] OF BOOL;(*横向启动延时标志*)
	axHorzMotorStart_DelayDne: ARRAY [1..MAX_UNIT_NUM] OF BOOL;(*横向启动延时完成*)
	auiHorzMotorStart_Count: ARRAY [1..MAX_UNIT_NUM] OF UINT;(*启动延时计时变量*)
	iHorzMotorStart_DelayTime_MS: INT:=0;(*启动的延时时间ms*)

	adwTotalTimes_CW_AxisHorzManu: ARRAY [1..MAX_UNIT_NUM] OF DWORD ;
	adwTotalTimes_CCW_AxisHorzManu: ARRAY [1..MAX_UNIT_NUM] OF DWORD ;
	lrAdjustVal_H_PerCycle:LREAL;(*每个周期调整的量*)

	(*2023.3.8.114227 将函数KS_FB_AxisHorAdj中的代码移植到此处*)
	axAxisHorAdjSts: ARRAY [1..MAX_UNIT_NUM] OF BOOL;
	axAxisHorAdj_End: ARRAY [1..MAX_UNIT_NUM] OF BOOL;
	iRtn: INT;
	iAdjustment_HorAxisAdj: INT;
	axHorAxisAdjStop: ARRAY [1..MAX_UNIT_NUM] OF BOOL;
	axHorAxisAdjStart: ARRAY [1..MAX_UNIT_NUM] OF BOOL;
	xFlag_HorAxisAdj: BOOL;
	wSts_HorzManuPreReg:WORD;
	(*横向运动相关变量都使用操作侧和传动侧变量重新赋值@2023.3.8.104853*)
	axHorMovingBtn_M: ARRAY [1..MAX_UNIT_NUM] OF BOOL;(*横向操作侧运动按钮*)
	axHorMovingBtn_G: ARRAY [1..MAX_UNIT_NUM] OF BOOL;(*横向传动侧运动按钮*)
	axHorMovingLimit_M: ARRAY [1..MAX_UNIT_NUM] OF BOOL;(*横向操作侧运动限位*)
	axHorMovingLimit_G: ARRAY [1..MAX_UNIT_NUM] OF BOOL;(*横向传动侧运动限位*)
	axHorMoving_M: ARRAY [1..MAX_UNIT_NUM] OF BOOL;(*横向操作侧运动*)
	axHorMoving_G: ARRAY [1..MAX_UNIT_NUM] OF BOOL;(*横向传动侧运动*)
	xAutoMove_H: BOOL;(*2025.4.20.110711+*)
END_VAR

{IMPLEMENTATION}
o_xEno:= i_xEn;
o_iErNo:= 0;
IF i_xEn THEN
	IF (i_iGrpAxisNum_Pu>=1 AND i_iGrpAxisNum_Pu<=MAX_UNIT_NUM) AND(*系的色组数量有效|*)
		i_pastStIOMap_AxisBasic<>0 AND
		i_pastStIOMap_AxisExtra<>0 THEN

		(*2023.3.8.114227 将函数KS_FB_AxisHorAdj中的代码移植到此处*)
		FOR iN:= 1 TO i_iGrpAxisNum_Pu BY 1 DO
			iUnitId:= i_abyGrpAxisList[iN];
			pstStIOMap_AxisBasic:= ADR(i_pastStIOMap_AxisBasic^[iUnitId]);

			(*处理横向开关相关@2023.3.8.104924*)
			(*和运动方向关联@伺服正转(正手机)-左对应操作侧#先不关心反印时候的方向变化问题
						    @伺服反转(反手机)-左对应传动侧#先不关心反印时候的方向变化问题*)
			IF NOT i_pstStSysParam^.astStUnitParam_UnSave[iUnitId].xMotRev_PrnRoller THEN(*正转*)
				axHorMovingBtn_M[iUnitId]:=pstStIOMap_AxisBasic^.i_xMove_Left;
				axHorMovingBtn_G[iUnitId]:=pstStIOMap_AxisBasic^.i_xMove_Right;

				axHorMovingLimit_M[iUnitId]:=pstStIOMap_AxisBasic^.i_xPosLimit_Left;
				axHorMovingLimit_G[iUnitId]:=pstStIOMap_AxisBasic^.i_xPosLimit_Right;
			ELSE(*反转*)
				axHorMovingBtn_M[iUnitId]:=pstStIOMap_AxisBasic^.i_xMove_Right;
				axHorMovingBtn_G[iUnitId]:=pstStIOMap_AxisBasic^.i_xMove_Left;

				IF i_xHorLimit THEN
					(*使用左右限位*)
					axHorMovingLimit_M[iUnitId]:=pstStIOMap_AxisBasic^.i_xPosLimit_Right;
					axHorMovingLimit_G[iUnitId]:=pstStIOMap_AxisBasic^.i_xPosLimit_Left;
				ELSE
					(*使用正转(操作侧)反转(传动侧)限位*)
					axHorMovingLimit_M[iUnitId]:=pstStIOMap_AxisBasic^.i_xPosLimit_Left;
					axHorMovingLimit_G[iUnitId]:=pstStIOMap_AxisBasic^.i_xPosLimit_Right;
				END_IF
			END_IF

			(*--------------------------------------------------|2019.11.18.153930_*)
			(*横向快速对版改成单个轴处理时放在循环内处理|*)
			(*返回的距离单位是mm*)
			iAdjustment_HorAxisAdj:=0;(*清零*)
			iRtn:= KS_FetchRapidAdjValue_H(i_pastStAxisRapidAdjProf_H, iUnitId, ADR(iAdjustment_HorAxisAdj));
			(*2024.01.17.161205 增加清除处理*)
			axHorAxisAdjStart[iUnitId]:= FALSE;
			axHorAxisAdjStop[iUnitId]:= FALSE;
			IF iRtn=0 THEN
				IF iAdjustment_HorAxisAdj=-32767 THEN(*人为停止标志|*)
					axHorAxisAdjStop[iUnitId]:= TRUE;
				ELSIF iAdjustment_HorAxisAdj<>0 THEN
					axHorAxisAdjStart[iUnitId]:= TRUE;
				END_IF
			END_IF

			IF (NOT i_xFlag_Estop) (*AND i_xFlag_Stop*) THEN(*非急停*)
				(*2025.4.20.105720 修改条件*)
				IF i_xFlag_Stop THEN(*不用限制单联动*)
					xAutoMove_H:=TRUE;
				ELSE(*非停机状态下|只有单动的可以*)
					xAutoMove_H:=NOT i_pstStSysParam^.astStUnitParam_Save[iUnitId].xLinkage;
				END_IF
				IF xAutoMove_H(*pstStAxisParam^.xLinkage *)THEN
					IF axHorAxisAdjStart[iUnitId] AND (NOT axAxisHorAdjSts[iUnitId]) THEN(*开始运行*)
						axAxisHorAdjSts[iUnitId]:= TRUE;
					END_IF

					IF (axHorAxisAdjStop[iUnitId] AND axAxisHorAdjSts[iUnitId]) OR(*停止运行*)
						axAxisHorAdj_End[iUnitId] THEN(*控制结束了就停止*)
						axAxisHorAdjSts[iUnitId]:= FALSE;
					END_IF
				ELSE
					axAxisHorAdjSts[iUnitId]:= FALSE;
					IF i_pstStSysParam^.astStUnitParam_UnSave[iUnitId].alrTotalAdjustVal_ManuCoarse_vh[2]<>0 THEN
						i_pstStSysParam^.astStUnitParam_UnSave[iUnitId].alrTotalAdjustVal_ManuCoarse_vh[2]:= 0;
					END_IF

				END_IF
			ELSE
				IF axAxisHorAdjSts[iUnitId] THEN
					axAxisHorAdjSts[iUnitId]:= FALSE;(*急停或者非停机-直接停止运行*)
					i_pstStSysParam^.astStUnitParam_UnSave[iUnitId].alrTotalAdjustVal_ManuCoarse_vh[2]:= 0;
				END_IF
			END_IF

			IF pstStIOMap_AxisBasic^.o_xRel_Press OR (NOT pstStIOMap_AxisBasic^.i_xHorzMotor_FastSpd) THEN
			(*快调/慢调处理*)
				lrAdjustVal_H_PerCycle:= i_lrVel_HorzAdjust*INT_TO_LREAL(i_iCycleTime_Plc);
			ELSE
				lrAdjustVal_H_PerCycle:= i_lrVel_HorzPreRegister*INT_TO_LREAL(i_iCycleTime_Plc);
			END_IF

			IF axAxisHorAdjSts[iUnitId] THEN (*色组进入到横向对版状态*)
				xFlag_HorAxisAdj:= TRUE;

				(*2025.4.20.105821 屏蔽联动条件*)
				IF i_pstStSysParam^.astStUnitParam_Save[iUnitId].xLinkage OR TRUE THEN(*色组联动*)
					IF NOT axAxisHorAdj_End[iUnitId] THEN
						IF NOT o_axAxisHorAdjing[iUnitId] THEN
							o_axAxisHorAdjing[iUnitId]:= TRUE;
							(*横向对版量叠加到横向手动粗调仓库*)
							(*iAdjustment_HorAxisAdj正值需要往传动侧运动*)
							(*iAdjustment_HorAxisAdj 单位mm
							  alrTotalAdjustVal_ManuCoarse_vh[2] 单位um*)
							i_pstStSysParam^.astStUnitParam_UnSave[iUnitId].alrTotalAdjustVal_ManuCoarse_vh[2]:= i_pstStSysParam^.astStUnitParam_UnSave[iUnitId].alrTotalAdjustVal_ManuCoarse_vh[2]+iAdjustment_HorAxisAdj*1000;(*单位um*)
							(*alrTotalAdjustVal_ManuCoarse_vh[2] 负值是向传动侧运动的@故取反*)
							i_pstStSysParam^.astStUnitParam_UnSave[iUnitId].alrTotalAdjustVal_ManuCoarse_vh[2]:=-i_pstStSysParam^.astStUnitParam_UnSave[iUnitId].alrTotalAdjustVal_ManuCoarse_vh[2];
						ELSE

							IF (axHorMovingLimit_G[iUnitId] AND i_pstStSysParam^.astStUnitParam_UnSave[iUnitId].alrTotalAdjustVal_ManuCoarse_vh[2]<0) OR
								(axHorMovingLimit_M[iUnitId] AND i_pstStSysParam^.astStUnitParam_UnSave[iUnitId].alrTotalAdjustVal_ManuCoarse_vh[2]>0) THEN
								i_pstStSysParam^.astStUnitParam_UnSave[iUnitId].alrTotalAdjustVal_ManuCoarse_vh[2]:=0;
							END_IF

							IF i_pstStSysParam^.astStUnitParam_UnSave[iUnitId].alrTotalAdjustVal_ManuCoarse_vh[2]=0 THEN(*调整量消耗完成*)
								o_axAxisHorAdjing[iUnitId]:= FALSE;
								axAxisHorAdj_End[iUnitId]:= TRUE;
							END_IF
						END_IF
					END_IF
				ELSE(*单动*)
					o_axAxisHorAdjing[iUnitId]:= FALSE;
					axAxisHorAdj_End[iUnitId]:= TRUE;
					IF i_pstStSysParam^.astStUnitParam_UnSave[iUnitId].alrTotalAdjustVal_ManuCoarse_vh[2]<>0 THEN
						i_pstStSysParam^.astStUnitParam_UnSave[iUnitId].alrTotalAdjustVal_ManuCoarse_vh[2]:=0;
					END_IF
				END_IF
			ELSE
				IF xFlag_HorAxisAdj THEN
					xFlag_HorAxisAdj:= FALSE;
				END_IF
				o_axAxisHorAdjing[iUnitId]:= FALSE;
				axAxisHorAdj_End[iUnitId]:= FALSE;
				IF i_pstStSysParam^.astStUnitParam_UnSave[iUnitId].alrTotalAdjustVal_ManuCoarse_vh[2]<>0 THEN(*退出横向对版状态，调整量清零*)
					i_pstStSysParam^.astStUnitParam_UnSave[iUnitId].alrTotalAdjustVal_ManuCoarse_vh[2]:=0;
				END_IF
			END_IF

			IF axAxisHorAdjSts[iUnitId] THEN
				IF ABS(i_pstStSysParam^.astStUnitParam_UnSave[iUnitId].alrTotalAdjustVal_ManuCoarse_vh[2])>=lrAdjustVal_H_PerCycle THEN
					IF i_pstStSysParam^.astStUnitParam_UnSave[iUnitId].alrTotalAdjustVal_ManuCoarse_vh[2]>0 THEN
						(*正向*)
						i_pstStSysParam^.astStUnitParam_UnSave[iUnitId].alrCurCycleAdjustVal_ManuCoarse_vh[2]:= lrAdjustVal_H_PerCycle;
						i_pstStSysParam^.astStUnitParam_UnSave[iUnitId].alrTotalAdjustVal_ManuCoarse_vh[2]:= i_pstStSysParam^.astStUnitParam_UnSave[iUnitId].alrTotalAdjustVal_ManuCoarse_vh[2] - i_pstStSysParam^.astStUnitParam_UnSave[iUnitId].alrCurCycleAdjustVal_ManuCoarse_vh[2];
						i_pstStSysParam^.astStUnitParam_UnSave[iUnitId].axCurCycleAdjustVal_ManuCoarse_done_vh[2]:= FALSE;
						axHorMovingBtn_M[iUnitId]:=TRUE;
						axHorMovingBtn_G[iUnitId]:=FALSE;
					ELSE
						(*反向*)
						i_pstStSysParam^.astStUnitParam_UnSave[iUnitId].alrCurCycleAdjustVal_ManuCoarse_vh[2]:= -lrAdjustVal_H_PerCycle;
						i_pstStSysParam^.astStUnitParam_UnSave[iUnitId].alrTotalAdjustVal_ManuCoarse_vh[2]:= i_pstStSysParam^.astStUnitParam_UnSave[iUnitId].alrTotalAdjustVal_ManuCoarse_vh[2] - i_pstStSysParam^.astStUnitParam_UnSave[iUnitId].alrCurCycleAdjustVal_ManuCoarse_vh[2];
						i_pstStSysParam^.astStUnitParam_UnSave[iUnitId].axCurCycleAdjustVal_ManuCoarse_done_vh[2]:= FALSE;

						axHorMovingBtn_M[iUnitId]:=FALSE;
						axHorMovingBtn_G[iUnitId]:=TRUE;
					END_IF
				ELSE
					IF o_axAxisHorAdjing[iUnitId] THEN
						i_pstStSysParam^.astStUnitParam_UnSave[iUnitId].alrTotalAdjustVal_ManuCoarse_vh[2]:= 0;
					END_IF
				END_IF
			END_IF
	(*往从站发送*)
			i_pstStSysParam^.astStUnitParam_UnSave[iUnitId].iPos_HorzManuPreReg:= -LREAL_TO_INT(i_pstStSysParam^.astStUnitParam_UnSave[iUnitId].alrTotalAdjustVal_ManuCoarse_vh[2]/1000);
			(*2024.01.17.170711 替换*)
			wSts_HorzManuPreReg.0:= axAxisHorAdjSts[iUnitId](*o_axAxisHorAdjing[iUnitId]*);
			wSts_HorzManuPreReg.1:= axHorMoving_M[iUnitId];
			wSts_HorzManuPreReg.2:= axHorMoving_G[iUnitId];
			wSts_HorzManuPreReg.3:= axHorMovingLimit_M[iUnitId];
			wSts_HorzManuPreReg.4:= axHorMovingLimit_G[iUnitId];
			wSts_HorzManuPreReg.5:= i_pstStSysParam^.astStGrpParam_UnSave[i_iGrpId].xFlag_Stop;

			i_pstStSysParam^.astStUnitParam_UnSave[iUnitId].wSts_HorzManuPreReg:= wSts_HorzManuPreReg;
		END_FOR

		IF i_pstStSysParam^.astStGrpParam_UnSave[i_iGrpId].xSts_HorzPreRegister THEN (*横向预套准状态*)
			xFlag_PreRegister_H:=TRUE;
			FOR iN:=1 TO i_iGrpAxisNum_Pu BY 1 DO
(*2019.03.15.142555|niu.j|放在IF外*)
				iUnitId:= i_abyGrpAxisList[iN];
				pstStIOMap_AxisBasic:= ADR(i_pastStIOMap_AxisBasic^[iUnitId]);
				pstStIOMap_AxisExtra:= ADR(i_pastStIOMap_AxisExtra^[iUnitId]);

				IF pstStIOMap_AxisBasic^.o_xRel_Press OR (NOT pstStIOMap_AxisBasic^.i_xHorzMotor_FastSpd) THEN
				(*快调/慢调处理*)
					lrAdjustVal_H_PerCycle:= i_lrVel_HorzAdjust*INT_TO_LREAL(i_iCycleTime_Plc);
				ELSE
					lrAdjustVal_H_PerCycle:= i_lrVel_HorzPreRegister*INT_TO_LREAL(i_iCycleTime_Plc);
				END_IF

				IF NOT 	i_pstStSysParam^.astStGrpParam_UnSave[i_iGrpId].xMode_HorzPreRegister THEN (*false 代表设定值 ，true代表重复值*)(*设定值！！走到左限位以目标值+当前修正量的值*)

					IF i_pstStSysParam^.astStUnitParam_Save[iUnitId].xLinkage THEN (*当前色处于联动状态才进行横向预套准*)
						IF NOT i_pstStSysParam^.astStUnitParam_UnSave[iUnitId].xFlag_HorzPreRegister_end THEN (*未调整完*)
							IF NOT i_pstStSysParam^.astStUnitParam_UnSave[iUnitId].xFlag_HorzPreRegister_ing THEN (*非横向预套准中*)
								IF NOT axHorMovingLimit_M[iUnitId] THEN (*未到操作侧限位*)
									i_pstStSysParam^.astStUnitParam_UnSave[iUnitId].alrTotalAdjustVal_Auto_vh[2]:=(2*lrAdjustVal_H_PerCycle);(*为了电机向左一直转动 diHorAdjValue_Sum>0,并且让他=一个周期调整的量*)

								ELSE(*到了操作侧限位*)
									i_pstStSysParam^.astStUnitParam_UnSave[iUnitId].xFlag_HorzPreRegister_ing:=TRUE;
									(*调整量单位um*)
									(*需要向传动侧运动*)
									i_pstStSysParam^.astStUnitParam_UnSave[iUnitId].alrTotalAdjustVal_Auto_vh[2]:=dint_to_lreal(i_pstStSysParam^.astStUnitParam_UnSave[iUnitId].diPreReg_SetupVal_H)*1000.0(*.diHorzPreReg_SetupVal*)+dint_to_lreal(i_pstStSysParam^.astStUnitParam_Save[iUnitId].diPreReg_AdjustVal_H)*1000.0(*.diHorzPreReg_AdjustVal*);(*设定值+修正值*)
									IF i_pstStSysParam^.astStUnitParam_UnSave[iUnitId].alrTotalAdjustVal_Auto_vh[2]<0 THEN
										i_pstStSysParam^.astStUnitParam_UnSave[iUnitId].alrTotalAdjustVal_Auto_vh[2]:=0;
									END_IF
									(*位置值为负值才是向传动侧运动的*)
									i_pstStSysParam^.astStUnitParam_UnSave[iUnitId].alrTotalAdjustVal_Auto_vh[2]:=-i_pstStSysParam^.astStUnitParam_UnSave[iUnitId].alrTotalAdjustVal_Auto_vh[2];
								END_IF
							ELSE(*预套准中*)
								IF axHorMovingLimit_G[iUnitId] THEN (*到达了传动侧限位*)
									i_pstStSysParam^.astStUnitParam_UnSave[iUnitId].alrTotalAdjustVal_Auto_vh[2]:=0;
								END_IF

								IF i_pstStSysParam^.astStUnitParam_UnSave[iUnitId].alrTotalAdjustVal_Auto_vh[2] =0 THEN(*预套准走完了*)
									i_pstStSysParam^.astStUnitParam_UnSave[iUnitId].xFlag_HorzPreRegister_ing:=FALSE;
									i_pstStSysParam^.astStUnitParam_UnSave[iUnitId].xFlag_HorzPreRegister_end:=TRUE;
								END_IF
							END_IF
						END_IF
					ELSE(*单动中*)
						i_pstStSysParam^.astStUnitParam_UnSave[iUnitId].xFlag_HorzPreRegister_ing:=FALSE;
						i_pstStSysParam^.astStUnitParam_UnSave[iUnitId].xFlag_HorzPreRegister_end:=TRUE;
						IF i_pstStSysParam^.astStUnitParam_UnSave[iUnitId].alrTotalAdjustVal_Auto_vh[2]<>0 THEN
							i_pstStSysParam^.astStUnitParam_UnSave[iUnitId].alrTotalAdjustVal_Auto_vh[2]:=0;
						END_IF
					END_IF

				ELSE(*重复值*)
					IF i_pstStSysParam^.astStUnitParam_Save[iUnitId].xLinkage THEN (*当前色处于联动状态才进行横向预套准*)
						IF NOT i_pstStSysParam^.astStUnitParam_UnSave[iUnitId].xFlag_HorzPreRegister_end THEN (*未调整完*)
							IF NOT i_pstStSysParam^.astStUnitParam_UnSave[iUnitId].xFlag_HorzPreRegister_ing THEN (*非横向预套准中*)
								i_pstStSysParam^.astStUnitParam_UnSave[iUnitId].xFlag_HorzPreRegister_ing:=TRUE;
								(*diPreReg_RepeatVal_H 正值向传动侧运动
								alrTotalAdjustVal_Auto_vh[2] 负值才是向传动侧运动@故需要取反*)
								i_pstStSysParam^.astStUnitParam_UnSave[iUnitId].alrTotalAdjustVal_Auto_vh[2]:=-DINT_TO_LREAL(i_pstStSysParam^.astStUnitParam_UnSave[iUnitId].diPreReg_RepeatVal_H)*1000.0(*.diHorzPreReg_RepeatVal*);(*diHorzPreReg_RepeatVal为正值代表要向右转动*)
																			(*下面执行的时候 只有总的调整量小于0才会输出向右转信号，故取反*)

							ELSE(*预套准中*)
								IF (axHorMovingLimit_G[iUnitId] AND i_pstStSysParam^.astStUnitParam_UnSave[iUnitId].alrTotalAdjustVal_Auto_vh[2]<0) OR
									(axHorMovingLimit_M[iUnitId] AND i_pstStSysParam^.astStUnitParam_UnSave[iUnitId].alrTotalAdjustVal_Auto_vh[2]>0) THEN
									i_pstStSysParam^.astStUnitParam_UnSave[iUnitId].alrTotalAdjustVal_Auto_vh[2]:=0;
								END_IF

								IF i_pstStSysParam^.astStUnitParam_UnSave[iUnitId].alrTotalAdjustVal_Auto_vh[2] =0 THEN(*预套准走完了*)
									i_pstStSysParam^.astStUnitParam_UnSave[iUnitId].xFlag_HorzPreRegister_ing:=FALSE;
									i_pstStSysParam^.astStUnitParam_UnSave[iUnitId].xFlag_HorzPreRegister_end:=TRUE;
								END_IF
							END_IF
						END_IF
					ELSE(*单动中*)
						i_pstStSysParam^.astStUnitParam_UnSave[iUnitId].xFlag_HorzPreRegister_ing:=FALSE;
						i_pstStSysParam^.astStUnitParam_UnSave[iUnitId].xFlag_HorzPreRegister_end:=TRUE;
						IF i_pstStSysParam^.astStUnitParam_UnSave[iUnitId].alrTotalAdjustVal_Auto_vh[2]<>0 THEN
							i_pstStSysParam^.astStUnitParam_UnSave[iUnitId].alrTotalAdjustVal_Auto_vh[2]:=0;
						END_IF
					END_IF
				END_IF
			END_FOR

			FOR iN:=1 TO i_iGrpAxisNum_Pu BY 1 DO(*检查所有的色组是否都完成*)
				iUnitId:= i_abyGrpAxisList[iN];

				IF i_pstStSysParam^.astStUnitParam_UnSave[iUnitId].xFlag_HorzPreRegister_end THEN
					i_pstStSysParam^.astStGrpParam_UnSave[i_iGrpId].xFlag_HorzPreRegister_All_end :=TRUE;(*横向预套准完成了*)
				ELSE
					i_pstStSysParam^.astStGrpParam_UnSave[i_iGrpId].xFlag_HorzPreRegister_All_end:=FALSE;
					EXIT;
				END_IF
			END_FOR

		ELSE(*非横向预套准中*)
			FOR iN:=1 TO i_iGrpAxisNum_Pu BY 1 DO(*检查所有的色组是否都完成*)
				iUnitId:= i_abyGrpAxisList[iN];

				i_pstStSysParam^.astStUnitParam_UnSave[iUnitId].xFlag_HorzPreRegister_ing:=FALSE;
				i_pstStSysParam^.astStUnitParam_UnSave[iUnitId].xFlag_HorzPreRegister_end:=FALSE;
			END_FOR

			IF xFlag_PreRegister_H THEN
				xFlag_PreRegister_H:=FALSE;
				FOR iN:=1 TO i_iGrpAxisNum_Pu BY 1 DO(*检查所有的色组是否都完成*)
					iUnitId:= i_abyGrpAxisList[iN];

					i_pstStSysParam^.astStUnitParam_UnSave[iUnitId].alrTotalAdjustVal_Auto_vh[2]:=0;
				END_FOR
			END_IF
			i_pstStSysParam^.astStGrpParam_UnSave[i_iGrpId].xFlag_HorzPreRegister_All_end:=FALSE;
		END_IF

		FOR iN:=1 TO i_iGrpAxisNum_Pu BY 1 DO
			iUnitId:= i_abyGrpAxisList[iN];
			pstStIOMap_AxisBasic:= ADR(i_pastStIOMap_AxisBasic^[iUnitId]);
			pstStIOMap_AxisExtra:= ADR(i_pastStIOMap_AxisExtra^[iUnitId]);

			IF pstStIOMap_AxisBasic^.o_xRel_Press OR (NOT pstStIOMap_AxisBasic^.i_xHorzMotor_FastSpd) THEN
			(*快调/慢调处理*)
				lrAdjustVal_H_PerCycle:= i_lrVel_HorzAdjust*INT_TO_LREAL(i_iCycleTime_Plc);
			ELSE
				lrAdjustVal_H_PerCycle:= i_lrVel_HorzPreRegister*INT_TO_LREAL(i_iCycleTime_Plc);
			END_IF

			(*2019.5.15.170941|niu.j|急停清零横向调整量*)
			IF i_pstStSysParam^.astStGrpParam_UnSave[i_iGrpId].xFlag_EStoping OR i_pstStSysParam^.astStGrpParam_UnSave[i_iGrpId].xFlag_Estop THEN
				i_pstStSysParam^.astStUnitParam_UnSave[iUnitId].alrTotalAdjustVal_Auto_vh[2]:= 0;
				i_pstStSysParam^.astStUnitParam_UnSave[iUnitId].alrTotalAdjustVal_ManuFine_vh[2]:= 0;
				i_pstStSysParam^.astStUnitParam_UnSave[iUnitId].alrTotalAdjustVal_Rapid_vh[2]:= 0;
			END_IF

			IF (i_pstStSysParam^.astStUnitParam_Save[iUnitId].dwFlag_Ctl.0 AND i_pstStSysParam^.astStUnitParam_Save[iUnitId].dwFlag_Sts.1)
				OR i_pstStSysParam^.astStGrpParam_UnSave[i_iGrpId].xSts_HorzPreRegister  THEN(*横向开|横向自动|*)
				(*消耗自动调整量累计|*)
				IF ABS(i_pstStSysParam^.astStUnitParam_UnSave[iUnitId].alrTotalAdjustVal_Auto_vh[2])>=lrAdjustVal_H_PerCycle THEN
					IF i_pstStSysParam^.astStUnitParam_UnSave[iUnitId].alrTotalAdjustVal_Auto_vh[2]>0 THEN
						(*正向*)
						i_pstStSysParam^.astStUnitParam_UnSave[iUnitId].alrCurCycleAdjustVal_Auto_vh[2]:= lrAdjustVal_H_PerCycle;
						i_pstStSysParam^.astStUnitParam_UnSave[iUnitId].alrTotalAdjustVal_Auto_vh[2]:= i_pstStSysParam^.astStUnitParam_UnSave[iUnitId].alrTotalAdjustVal_Auto_vh[2] - i_pstStSysParam^.astStUnitParam_UnSave[iUnitId].alrCurCycleAdjustVal_Auto_vh[2];
						i_pstStSysParam^.astStUnitParam_UnSave[iUnitId].axCurCycleAdjustVal_Auto_done_vh[2]:= FALSE;
						axHorMoving_M[iUnitId]:= TRUE;(*操作侧*)
						axHorMoving_G[iUnitId]:= FALSE;(*传动侧*)
					ELSE
						(*反向*)
						i_pstStSysParam^.astStUnitParam_UnSave[iUnitId].alrCurCycleAdjustVal_Auto_vh[2]:= -lrAdjustVal_H_PerCycle;
						i_pstStSysParam^.astStUnitParam_UnSave[iUnitId].alrTotalAdjustVal_Auto_vh[2]:= i_pstStSysParam^.astStUnitParam_UnSave[iUnitId].alrTotalAdjustVal_Auto_vh[2] - i_pstStSysParam^.astStUnitParam_UnSave[iUnitId].alrCurCycleAdjustVal_Auto_vh[2];
						i_pstStSysParam^.astStUnitParam_UnSave[iUnitId].axCurCycleAdjustVal_Auto_done_vh[2]:= FALSE;
						axHorMoving_G[iUnitId]:= TRUE;(*传动侧*)
						axHorMoving_M[iUnitId]:= FALSE;(*操作侧*)
					END_IF
				ELSE
					IF i_pstStSysParam^.astStUnitParam_UnSave[iUnitId].xFlag_HorzPreRegister_ing THEN
						i_pstStSysParam^.astStUnitParam_UnSave[iUnitId].alrTotalAdjustVal_Auto_vh[2]:= 0;
					END_IF
					//2025.9.9.200410 同步
					(*2025.9.5.104621 对于小调整量进行响应处理优化*)
					IF lrAdjustVal_H_PerCycle > 10 THEN(*单周期的量超过1丝执行这部分代码*)
						IF ABS(i_pstStSysParam^.astStUnitParam_UnSave[iUnitId].alrTotalAdjustVal_Auto_vh[2]) >= 10 THEN(*强制响应1丝以上的调整量*)
							IF i_pstStSysParam^.astStUnitParam_UnSave[iUnitId].alrTotalAdjustVal_Auto_vh[2] > 0 THEN(*正向*)
								axHorMoving_M[iUnitId]:= TRUE;(*操作侧*)
								axHorMoving_G[iUnitId]:= FALSE;(*传动侧*)
							ELSE(*反向*)
								axHorMoving_M[iUnitId]:= FALSE;(*操作侧*)
								axHorMoving_G[iUnitId]:= TRUE;(*传动侧*)
							END_IF
							i_pstStSysParam^.astStUnitParam_UnSave[iUnitId].alrTotalAdjustVal_Auto_vh[2]:=0;(*清零*)
						ELSE
							axHorMoving_M[iUnitId]:= FALSE;(*操作侧*)
							axHorMoving_G[iUnitId]:= FALSE;(*传动侧*)
						END_IF
					ELSE(*单周期的量小于1丝的时候就不响应剩余的调整量*)
						axHorMoving_M[iUnitId]:= FALSE;(*操作侧*)
						axHorMoving_G[iUnitId]:= FALSE;(*传动侧*)
					END_IF
				END_IF
			ELSIF i_xHorManuCtrl THEN(*界面上有横向手动修正功能|*)
				(*消耗手动细调量累计|*)
				IF ABS(i_pstStSysParam^.astStUnitParam_UnSave[iUnitId].alrTotalAdjustVal_ManuFine_vh[2])>=lrAdjustVal_H_PerCycle THEN
(*					IF axHorzMotorStart_DelayDne[iUnitId] THEN(*延时启动完成了*)
*)						IF i_pstStSysParam^.astStUnitParam_UnSave[iUnitId].alrTotalAdjustVal_ManuFine_vh[2]>0 THEN
							(*正向*)
							i_pstStSysParam^.astStUnitParam_UnSave[iUnitId].alrCurCycleAdjustVal_ManuFine_vh[2]:= lrAdjustVal_H_PerCycle;

							i_pstStSysParam^.astStUnitParam_UnSave[iUnitId].alrTotalAdjustVal_ManuFine_vh[2]:= i_pstStSysParam^.astStUnitParam_UnSave[iUnitId].alrTotalAdjustVal_ManuFine_vh[2] - i_pstStSysParam^.astStUnitParam_UnSave[iUnitId].alrCurCycleAdjustVal_ManuFine_vh[2];
							i_pstStSysParam^.astStUnitParam_UnSave[iUnitId].axCurCycleAdjustVal_ManuFine_done_vh[2]:= FALSE;
							axHorMoving_M[iUnitId]:= TRUE;(*操作侧*)
							axHorMoving_G[iUnitId]:= FALSE;(*传动侧*)

						ELSE
							(*反向*)
							i_pstStSysParam^.astStUnitParam_UnSave[iUnitId].alrCurCycleAdjustVal_ManuFine_vh[2]:= -lrAdjustVal_H_PerCycle;

							i_pstStSysParam^.astStUnitParam_UnSave[iUnitId].alrTotalAdjustVal_ManuFine_vh[2]:= i_pstStSysParam^.astStUnitParam_UnSave[iUnitId].alrTotalAdjustVal_ManuFine_vh[2] - i_pstStSysParam^.astStUnitParam_UnSave[iUnitId].alrCurCycleAdjustVal_ManuFine_vh[2];
							i_pstStSysParam^.astStUnitParam_UnSave[iUnitId].axCurCycleAdjustVal_ManuFine_done_vh[2]:= FALSE;
							axHorMoving_G[iUnitId]:= TRUE;(*传动侧*)
							axHorMoving_M[iUnitId]:= FALSE;(*操作侧*)

						END_IF

					(*monitoring...\2018.10.7.104410|*)
					IF axHorMoving_M[iUnitId] THEN
						adwTotalTimes_CW_AxisHorzManu[iUnitId]:= adwTotalTimes_CW_AxisHorzManu[iUnitId]+1;
					END_IF
					IF axHorMoving_G[iUnitId] THEN
						adwTotalTimes_CCW_AxisHorzManu[iUnitId]:= adwTotalTimes_CCW_AxisHorzManu[iUnitId]+1;
					END_IF

				ELSE

					axHorMoving_M[iUnitId]:= FALSE;
					axHorMoving_G[iUnitId]:= FALSE;
				END_IF
			ELSE
				(*没开横向或者横向在手动状态*)
				i_pstStSysParam^.astStUnitParam_UnSave[iUnitId].axCurCycleAdjustVal_Auto_done_vh[2]:= FALSE;
				i_pstStSysParam^.astStUnitParam_UnSave[iUnitId].axCurCycleAdjustVal_Rapid_done_vh[2]:= FALSE;
				i_pstStSysParam^.astStUnitParam_UnSave[iUnitId].axCurCycleAdjustVal_ManuCoarse_done_vh[2]:= FALSE;
				i_pstStSysParam^.astStUnitParam_UnSave[iUnitId].axCurCycleAdjustVal_ManuFine_done_vh[2]:= FALSE;
				i_pstStSysParam^.astStUnitParam_UnSave[iUnitId].axCurCycleAdjustVal_Coupling_done_vh[2]:= FALSE;
				i_pstStSysParam^.astStUnitParam_UnSave[iUnitId].axCurCycleAdjustVal_Compensate_done_vh[2]:= FALSE;

				i_pstStSysParam^.astStUnitParam_UnSave[iUnitId].alrCurCycleAdjustVal_Auto_vh[2]:= 0;
				i_pstStSysParam^.astStUnitParam_UnSave[iUnitId].alrCurCycleAdjustVal_Rapid_vh[2]:= 0;
				i_pstStSysParam^.astStUnitParam_UnSave[iUnitId].alrCurCycleAdjustVal_ManuCoarse_vh[2]:= 0;
				i_pstStSysParam^.astStUnitParam_UnSave[iUnitId].alrCurCycleAdjustVal_ManuFine_vh[2]:= 0;
				i_pstStSysParam^.astStUnitParam_UnSave[iUnitId].alrCurCycleAdjustVal_Coupling_vh[2]:= 0;
				i_pstStSysParam^.astStUnitParam_UnSave[iUnitId].alrCurCycleAdjustVal_Compensate_vh[2]:= 0;

				i_pstStSysParam^.astStUnitParam_UnSave[iUnitId].alrTotalAdjustVal_Auto_vh[2]:= 0;
				i_pstStSysParam^.astStUnitParam_UnSave[iUnitId].alrTotalAdjustVal_Rapid_vh[2]:= 0;
(*				pstStAxisParam^.alrTotalAdjustVal_ManuCoarse_vh[2]:= 0;*)
				i_pstStSysParam^.astStUnitParam_UnSave[iUnitId].alrTotalAdjustVal_ManuFine_vh[2]:= 0;
				i_pstStSysParam^.astStUnitParam_UnSave[iUnitId].alrTotalAdjustVal_Coupling_vh[2]:= 0;
				i_pstStSysParam^.astStUnitParam_UnSave[iUnitId].alrTotalAdjustVal_Compensate_vh[2]:= 0;

				axHorMoving_M[iUnitId]:= FALSE;
				axHorMoving_G[iUnitId]:= FALSE;
			END_IF
(*
			axHorzMotorStart_Delay[1];
			axHorzMotorStart_Delay[2];
			axHorzMotorStart_Delay[3];
			axHorzMotorStart_Delay[4];
			axHorzMotorStart_Delay[5];
			axHorzMotorStart_Delay[6];
			axHorzMotorStart_Delay[7];
			axHorzMotorStart_Delay[8];
			axHorzMotorStart_Delay[9];

			axHorzMotorStart_DelayDne[1];
			axHorzMotorStart_DelayDne[2];
			axHorzMotorStart_DelayDne[3];
			axHorzMotorStart_DelayDne[4];
			axHorzMotorStart_DelayDne[5];
			axHorzMotorStart_DelayDne[6];
			axHorzMotorStart_DelayDne[7];
			axHorzMotorStart_DelayDne[8];
			axHorzMotorStart_DelayDne[9];

			auiHorzMotorStart_Count[1];
			auiHorzMotorStart_Count[2];
			auiHorzMotorStart_Count[3];
			auiHorzMotorStart_Count[4];
			auiHorzMotorStart_Count[5];
			auiHorzMotorStart_Count[6];
			auiHorzMotorStart_Count[7];
			auiHorzMotorStart_Count[8];
			auiHorzMotorStart_Count[9];

			awPreHorzMotorDir[1];
			awPreHorzMotorDir[2];
			awPreHorzMotorDir[3];
			awPreHorzMotorDir[4];
			awPreHorzMotorDir[5];
			awPreHorzMotorDir[6];
			awPreHorzMotorDir[7];
			awPreHorzMotorDir[8];
			awPreHorzMotorDir[9];
*)

			(*增加了正反转信号启动延时2018.10.7.085705 by liu.yt*)
			wHorzMotorDir:=BOOL_TO_WORD(axHorMoving_M[iUnitId])+SHL(BOOL_TO_WORD(axHorMoving_G[iUnitId]),1);
			IF wHorzMotorDir<>awPreHorzMotorDir[iUnitId] THEN(*方向发生了变化*)
				IF wHorzMotorDir<>0THEN(*说明有正反转信号了*)
					axHorzMotorStart_Delay[iUnitId]:=TRUE;
				ELSE
					axHorzMotorStart_Delay[iUnitId]:=FALSE;
				END_IF
				axHorzMotorStart_DelayDne[iUnitId]:=FALSE;
				auiHorzMotorStart_Count[iUnitId]:=0;
				awPreHorzMotorDir[iUnitId]:=wHorzMotorDir;
			END_IF

			IF axHorzMotorStart_Delay[iUnitId] THEN(*启动延时*)
				IF auiHorzMotorStart_Count[iUnitId]>=iHorzMotorStart_DelayTime_MS/i_iCycleTime_Plc THEN
					auiHorzMotorStart_Count[iUnitId]:=0;
					axHorzMotorStart_Delay[iUnitId]:=FALSE;
					axHorzMotorStart_DelayDne[iUnitId]:=TRUE;
				ELSE
					auiHorzMotorStart_Count[iUnitId]:=auiHorzMotorStart_Count[iUnitId]+1;
				END_IF
			END_IF

			(*---------------------------2017-08-14 15:21:18
			/.手动调整
			.----------------------------------------------*)
			IF axHorMovingBtn_M[iUnitId] AND (NOT axHorMovingBtn_G[iUnitId]) THEN
				(*左*)
				axHorMoving_G[iUnitId]:= FALSE;
				axHorMoving_M[iUnitId]:= TRUE;
			ELSIF axHorMovingBtn_G[iUnitId] AND (NOT axHorMovingBtn_M[iUnitId]) THEN
				(*右*)
				axHorMoving_M[iUnitId]:= FALSE;
				axHorMoving_G[iUnitId]:= TRUE;
			END_IF

			(*---------------------------2017-08-14 15:21:18
			/.横向限位处理
			.----------------------------------------------*)
			IF axHorMovingLimit_M[iUnitId] THEN(*操作侧*)
				axHorMoving_M[iUnitId]:= FALSE;
			END_IF

			IF axHorMovingLimit_G[iUnitId] THEN(*传动侧*)
				axHorMoving_G[iUnitId]:= FALSE;
			END_IF

			(*急停停止横向输出|2022.5.11.171513*)
			IF i_pstStSysParam^.astStGrpParam_UnSave[i_iGrpId].xFlag_EStoping OR i_pstStSysParam^.astStGrpParam_UnSave[i_iGrpId].xFlag_Estop THEN
				axHorMoving_M[iUnitId]:= FALSE;
				axHorMoving_G[iUnitId]:= FALSE;
			END_IF

			(*将操作侧和传动侧信号输出*)
			(*电机输出是按照正转和反转@一般情况正反手机电机的旋转方向是一致的即,都是向操作侧或者都是向传动侧
			我们定义正传是向操作侧@反转是向传动侧*)
			pstStIOMap_AxisBasic^.o_xHorzMotor_CW:=axHorMoving_M[iUnitId];
			pstStIOMap_AxisBasic^.o_xHorzMotor_CCW:=axHorMoving_G[iUnitId];
		END_FOR
	ELSE
		o_iErNo:= -1;
	END_IF
END_IF

(* ---- KS_FB_GrpHorzAdjCtl_Driver.st ---- *)
(*@CES
Name=KS_FB_GrpHorzAdjCtl_Driver
Type=FunctionBlock
TypeGuid=6f9dac99-8de1-4efc-8465-68ac443b7d08
Guid=05f0aed7-3c56-4fbb-a93f-ecb252c274d1
HasDeclaration=True
HasImplementation=True
*)
{DECLARATION}
FUNCTION_BLOCK KS_FB_GrpHorzAdjCtl_Driver
VAR_INPUT
	i_xEn: BOOL;
	i_iGrpAxisNum_Pu: INT;
	i_aiStationList_Trap: ARRAY [1..MAX_STATION_NUM] OF INT;
	i_pastStIOMap_AxisBasic					: POINTER TO ARRAY [1..MAX_UNIT_NUM] OF StIOMap_Axis_FE; (*基础io|*)

END_VAR
VAR_OUTPUT
	o_xEn: BOOL;
	o_iErNo: INT;
END_VAR
VAR
	iN: INT;
	xInit: BOOL;
	iAxisId: INT;
	pstStIOMap_Axis_FLEXO: POINTER TO StIOMap_Axis_FLEXO;
	pstStUnitParam: POINTER TO StUnitParam;

	(*横向运动相关变量都使用操作侧和传动侧变量重新赋值@2023.3.8.104853*)
	axHorMovingBtn_M: ARRAY [1..MAX_UNIT_NUM] OF BOOL;(*横向操作侧运动按钮*)
	axHorMovingBtn_G: ARRAY [1..MAX_UNIT_NUM] OF BOOL;(*横向传动侧运动按钮*)
	axHorMovingLimit_M: ARRAY [1..MAX_UNIT_NUM] OF BOOL;(*横向操作侧运动限位*)
	axHorMovingLimit_G: ARRAY [1..MAX_UNIT_NUM] OF BOOL;(*横向传动侧运动限位*)
	axHorMoving_M: ARRAY [1..MAX_UNIT_NUM] OF BOOL;(*横向操作侧运动*)
	axHorMoving_G: ARRAY [1..MAX_UNIT_NUM] OF BOOL;(*横向传动侧运动*)

	lrAdjustVel_:LREAL;(*每个周期调整的量|这里还是mm/s，需要转化为*)
	alrTotalAdjust_Horz: ARRAY [1..MAX_UNIT_NUM] OF LREAL;(*横向调整量*)
	adwTotalTimes_CW_AxisHorzManu: ARRAY [1..MAX_UNIT_NUM] OF DWORD := [MAX_UNIT_NUM(0)];
	adwTotalTimes_CCW_AxisHorzManu: ARRAY [1..MAX_UNIT_NUM] OF DWORD := [MAX_UNIT_NUM(0)];

	wHorzMotorDir: WORD;(*.0 |正转方向
					.1|反转方向*)
	awPreHorzMotorDir: ARRAY [1..MAX_UNIT_NUM] OF WORD;
	axHorzMotorStart_Delay: ARRAY [1..MAX_UNIT_NUM] OF BOOL;(*横向启动延时标志*)
	axHorzMotorStart_DelayDne: ARRAY [1..MAX_UNIT_NUM] OF BOOL;(*横向启动延时完成*)
	auiHorzMotorStart_Count: ARRAY [1..MAX_UNIT_NUM] OF UINT;(*启动延时计时变量*)
	iHorzMotorStart_DelayTime_MS: INT:=0;(*启动的延时时间ms*)

	axStopManuMove_Horz: ARRAY  [1..MAX_UNIT_NUM] OF BOOL;
	lrLimit_Left:LREAL;
	lrLimit_Right:LREAL;
	xLimit_LeftTemp:BOOL;
	xLimit_RightTemp:BOOL;
	xLimit_Left:BOOL;
	xLimit_Right:BOOL;
END_VAR

{IMPLEMENTATION}
o_xEn:= i_xEn;
o_iErNo:= 0;
IF i_xEn THEN
	IF i_iGrpAxisNum_Pu>=1 AND i_iGrpAxisNum_Pu<=MAX_UNIT_NUM AND i_pastStIOMap_AxisBasic<>0 THEN
		IF NOT xInit THEN
			xInit:= TRUE;
			FOR iN:=1 TO i_iGrpAxisNum_Pu BY 1 DO
				alrTotalAdjust_Horz[iN]:= 0;
			END_FOR
		END_IF
		(*2023.3.8.114227 将函数KS_FB_AxisHorAdj中的代码移植到此处*)
		FOR iN:= 1 TO i_iGrpAxisNum_Pu BY 1 DO
			iAxisId:= iN;
			pstStUnitParam:= ADR(i_pstStSysParam^.astStUnitParam[iAxisId]);
			pstStIOMap_Axis_FLEXO:= ADR(i_pastStIOMap_Axis_FLEXO^[iAxisId]);

			(*处理一下限位*)
			(*限位赋值*)
			IF i_pstStSysParam^.xIsDebugMode_Machine AND i_pstStSysParam^.xFlag_Stop THEN//调试模式
				//记录一下横向限位
				IF i_paxLimit_Left_Wr^[iAxisId] THEN
					i_paxLimit_Left_Wr^[iAxisId]:= FALSE;
					pstStUnitParam^.lrLimit_Left:= i_alrTarp_EncPos[iAxisId];
				END_IF
				IF i_paxLimit_Right_Wr^[iAxisId] THEN
					i_paxLimit_Right_Wr^[iAxisId]:= FALSE;
					pstStUnitParam^.lrLimit_Right:= i_alrTarp_EncPos[iAxisId];
				END_IF
				IF 	i_paxLimit_Left_WrClr^[iAxisId] THEN
					i_paxLimit_Left_WrClr^[iAxisId] := FALSE;
					pstStUnitParam^.lrLimit_Left := 0;
				END_IF
				IF 	i_paxLimit_Right_WrClr^[iAxisId] THEN
					i_paxLimit_Right_WrClr^[iAxisId] := FALSE;
					pstStUnitParam^.lrLimit_Right := 0;
				END_IF
			ELSE
				i_paxLimit_Left_Wr^[iAxisId]:= FALSE;
				i_paxLimit_Right_Wr^[iAxisId]:= FALSE;
				i_paxLimit_Left_WrClr^[iAxisId]:= FALSE;
				i_paxLimit_Right_WrClr^[iAxisId]:= FALSE;
			END_IF
			lrLimit_Left:= pstStUnitParam^.lrLimit_Left;
			lrLimit_Right:= pstStUnitParam^.lrLimit_Right;
			xLimit_LeftTemp:=i_pastStIOMap_Axis_FLEXO^[iAxisId].i_xPosLimit_Left;
			xLimit_RightTemp:=i_pastStIOMap_Axis_FLEXO^[iAxisId].i_xPosLimit_Right;

			IF lrLimit_Left=0 THEN(*未有软限位|按照最远距离*);

			ELSE(*存在软限位|限位标志取接近开关和位置值的or*)
				IF pstStUnitParam^.xMotRev_Horiz_ THEN
					xLimit_LeftTemp:=xLimit_LeftTemp OR
									(lrLimit_Left<i_alrTarp_EncPos[iAxisId]);
				ELSE
					xLimit_LeftTemp:=xLimit_LeftTemp OR
									(lrLimit_Left>i_alrTarp_EncPos[iAxisId]);
				END_IF
			END_IF
			IF lrLimit_Right=0 THEN(*未有软限位|按照最远距离*);
			ELSE(*存在软限位|限位标志取接近开关和位置值的or*)
				IF pstStUnitParam^.xMotRev_Horiz_ THEN
					xLimit_RightTemp:=xLimit_RightTemp OR
								(lrLimit_Right>i_alrTarp_EncPos[iAxisId]);
				ELSE
					xLimit_RightTemp:=xLimit_RightTemp OR
								(lrLimit_Right<i_alrTarp_EncPos[iAxisId]);

				END_IF
			END_IF

			(*手动左右取反*)(*bai.zy|2023.12.18.161830|feida取反*)
			xLimit_Left:=xLimit_LeftTemp;
			xLimit_Right:=xLimit_RightTemp;
			IF pstStUnitParam^.xMotRev_Horiz_ THEN
				xLimit_Left:=xLimit_LeftTemp;
				xLimit_Right:=xLimit_RightTemp;
			END_IF
			g_axLimit_Left_Wr_HMI[iN]:= xLimit_Left;
			g_axLimit_Right_Wr_HMI[iN]:= xLimit_Right;
			(*处理横向开关相关@2023.3.8.104924*)
			(*和运动方向关联@伺服正转(正手机)-左对应操作侧#先不关心反印时候的方向变化问题
						    @伺服反转(反手机)-左对应传动侧#先不关心反印时候的方向变化问题*)

//			IF pstStUnitParam^.xMotRev_PrnRoller THEN(*正转*)
				axHorMovingBtn_M[iAxisId]:=pstStIOMap_Axis_FLEXO^.i_xMove_Left;
				axHorMovingBtn_G[iAxisId]:=pstStIOMap_Axis_FLEXO^.i_xMove_Right;

				axHorMovingLimit_M[iAxisId]:=xLimit_Left;
				axHorMovingLimit_G[iAxisId]:=xLimit_Right;
(*			ELSE(*反转*)
				axHorMovingBtn_M[iAxisId]:=pstStIOMap_Axis_FLEXO^.i_xMove_Right;
				axHorMovingBtn_G[iAxisId]:=pstStIOMap_Axis_FLEXO^.i_xMove_Left;

				IF i_pstStSysParam^.dwControlComplexBits.17 THEN
					(*使用左右限位*)
					axHorMovingLimit_M[iAxisId]:=xLimit_Right;
					axHorMovingLimit_G[iAxisId]:=xLimit_Left;
				ELSE
					(*使用正转(操作侧)反转(传动侧)限位*)
					axHorMovingLimit_M[iAxisId]:=xLimit_Left;
					axHorMovingLimit_G[iAxisId]:=xLimit_Right;
				END_IF
			END_IF
*)

			IF pstStIOMap_Axis_FLEXO^.o_xRel_Press OR (NOT pstStIOMap_Axis_FLEXO^.i_xHorzMotor_FastSpd) THEN
			(*快调/慢调处理*)
				lrAdjustVel_:= i_lrVel_HorzAdjust;
			ELSE
				lrAdjustVel_:= i_lrVel_HorzPreRegister;
			END_IF

			(*2019.5.15.170941|niu.j|急停清零横向调整量*)
			IF i_pstStSysParam^.xFlag_EStoping OR i_pstStSysParam^.xFlag_Estop THEN
				pstStUnitParam^.alrTotalAdjustVal_Auto_vh[2]:= 0;
				pstStUnitParam^.alrTotalAdjustVal_ManuFine_vh[2]:= 0;
				pstStUnitParam^.alrTotalAdjustVal_Rapid_vh[2]:= 0;
			END_IF

			IF (pstStUnitParam^.dwFlag_Ctl.0 AND pstStUnitParam^.dwFlag_Sts.1) THEN
				IF ABS(pstStUnitParam^.alrTotalAdjustVal_Auto_vh[2])>0 THEN
					IF pstStUnitParam^.alrTotalAdjustVal_Auto_vh[2]>0 THEN
						(*正向*)
						alrTotalAdjust_Horz[iAxisId]:= alrTotalAdjust_Horz[iAxisId]+pstStUnitParam^.alrTotalAdjustVal_Auto_vh[2];
						pstStUnitParam^.alrTotalAdjustVal_Auto_vh[2]:= 0;
						pstStUnitParam^.axCurCycleAdjustVal_Auto_done_vh[2]:= FALSE;
						axHorMoving_M[iAxisId]:= TRUE;(*操作侧*)
						axHorMoving_G[iAxisId]:= FALSE;(*传动侧*)
					ELSE
						(*反向*)
						alrTotalAdjust_Horz[iAxisId]:= alrTotalAdjust_Horz[iAxisId]+pstStUnitParam^.alrTotalAdjustVal_Auto_vh[2];
						pstStUnitParam^.alrTotalAdjustVal_Auto_vh[2]:= 0;
						pstStUnitParam^.axCurCycleAdjustVal_Auto_done_vh[2]:= FALSE;
						axHorMoving_G[iAxisId]:= TRUE;(*传动侧*)
						axHorMoving_M[iAxisId]:= FALSE;(*操作侧*)
					END_IF
				ELSE
					IF pstStUnitParam^.xFlag_HorzPreRegister_ing THEN
						pstStUnitParam^.alrTotalAdjustVal_Auto_vh[2]:= 0;
					END_IF
					axHorMoving_M[iAxisId]:= FALSE;
					axHorMoving_G[iAxisId]:= FALSE;
				END_IF
			ELSIF i_pstStSysParam^.dwControlComplexBits.7 THEN(*界面上有横向手动修正功能|*)
				(*消耗手动细调量累计|*)
				IF ABS(pstStUnitParam^.alrTotalAdjustVal_ManuFine_vh[2])>0 THEN
(*					IF axHorzMotorStart_DelayDne[iAxisId] THEN(*延时启动完成了*)
*)						IF pstStUnitParam^.alrTotalAdjustVal_ManuFine_vh[2]>0 THEN
							(*正向*)
							alrTotalAdjust_Horz[iAxisId]:= alrTotalAdjust_Horz[iAxisId]+pstStUnitParam^.alrTotalAdjustVal_ManuFine_vh[2];
							pstStUnitParam^.alrTotalAdjustVal_ManuFine_vh[2]:= 0;
							pstStUnitParam^.axCurCycleAdjustVal_ManuFine_done_vh[2]:= FALSE;
							axHorMoving_M[iAxisId]:= TRUE;(*操作侧*)
							axHorMoving_G[iAxisId]:= FALSE;(*传动侧*)

						ELSE
							(*反向*)
							alrTotalAdjust_Horz[iAxisId]:= alrTotalAdjust_Horz[iAxisId]+pstStUnitParam^.alrTotalAdjustVal_ManuFine_vh[2];
							pstStUnitParam^.alrTotalAdjustVal_ManuFine_vh[2]:= 0;
							pstStUnitParam^.axCurCycleAdjustVal_ManuFine_done_vh[2]:= FALSE;
							axHorMoving_G[iAxisId]:= TRUE;(*传动侧*)
							axHorMoving_M[iAxisId]:= FALSE;(*操作侧*)

						END_IF

					(*monitoring...\2018.10.7.104410|*)
					IF axHorMoving_M[iAxisId] THEN
						adwTotalTimes_CW_AxisHorzManu[iAxisId]:= adwTotalTimes_CW_AxisHorzManu[iAxisId]+1;
					END_IF
					IF axHorMoving_G[iAxisId] THEN
						adwTotalTimes_CCW_AxisHorzManu[iAxisId]:= adwTotalTimes_CCW_AxisHorzManu[iAxisId]+1;
					END_IF

				ELSE
					axHorMoving_M[iAxisId]:= FALSE;
					axHorMoving_G[iAxisId]:= FALSE;
				END_IF
			ELSE
				(*没开横向或者横向在手动状态*)
				pstStUnitParam^.axCurCycleAdjustVal_Auto_done_vh[2]:= FALSE;
				pstStUnitParam^.axCurCycleAdjustVal_Rapid_done_vh[2]:= FALSE;
				pstStUnitParam^.axCurCycleAdjustVal_ManuCoarse_done_vh[2]:= FALSE;
				pstStUnitParam^.axCurCycleAdjustVal_ManuFine_done_vh[2]:= FALSE;
				pstStUnitParam^.axCurCycleAdjustVal_Coupling_done_vh[2]:= FALSE;
//				pstStUnitParam^.axCurCycleAdjustVal_Compensate_done_vh[2]:= FALSE;

				pstStUnitParam^.alrCurCycleAdjustVal_Auto_vh[2]:= 0;
				pstStUnitParam^.alrCurCycleAdjustVal_Rapid_vh[2]:= 0;
				pstStUnitParam^.alrCurCycleAdjustVal_ManuCoarse_vh[2]:= 0;
				pstStUnitParam^.alrCurCycleAdjustVal_ManuFine_vh[2]:= 0;
				pstStUnitParam^.alrCurCycleAdjustVal_Coupling_vh[2]:= 0;
//				pstStUnitParam^.alrCurCycleAdjustVal_Compensate_vh[2]:= 0;

				pstStUnitParam^.alrTotalAdjustVal_Auto_vh[2]:= 0;
				pstStUnitParam^.alrTotalAdjustVal_Rapid_vh[2]:= 0;
(*				pstStUnitParam^.alrTotalAdjustVal_ManuCoarse_vh[2]:= 0;*)
				pstStUnitParam^.alrTotalAdjustVal_ManuFine_vh[2]:= 0;
				pstStUnitParam^.alrTotalAdjustVal_Coupling_vh[2]:= 0;
//				pstStUnitParam^.alrTotalAdjustVal_Compensate_vh[2]:= 0;

				axHorMoving_M[iAxisId]:= FALSE;
				axHorMoving_G[iAxisId]:= FALSE;
			END_IF

			(*增加了正反转信号启动延时2018.10.7.085705 by liu.yt*)
			wHorzMotorDir:=BOOL_TO_WORD(axHorMoving_M[iAxisId])+SHL(BOOL_TO_WORD(axHorMoving_G[iAxisId]),1);
			IF wHorzMotorDir<>awPreHorzMotorDir[iAxisId] THEN(*方向发生了变化*)
				IF wHorzMotorDir<>0THEN(*说明有正反转信号了*)
					axHorzMotorStart_Delay[iAxisId]:=TRUE;
				ELSE
					axHorzMotorStart_Delay[iAxisId]:=FALSE;
				END_IF
				axHorzMotorStart_DelayDne[iAxisId]:=FALSE;
				auiHorzMotorStart_Count[iAxisId]:=0;
				awPreHorzMotorDir[iAxisId]:=wHorzMotorDir;
			END_IF

			IF axHorzMotorStart_Delay[iAxisId] THEN(*启动延时*)
				IF auiHorzMotorStart_Count[iAxisId]>=iHorzMotorStart_DelayTime_MS/i_iCycleTime_Plc THEN
					auiHorzMotorStart_Count[iAxisId]:=0;
					axHorzMotorStart_Delay[iAxisId]:=FALSE;
					axHorzMotorStart_DelayDne[iAxisId]:=TRUE;
				ELSE
					auiHorzMotorStart_Count[iAxisId]:=auiHorzMotorStart_Count[iAxisId]+1;
				END_IF
			END_IF

			(*---------------------------2017-08-14 15:21:18
			/.手动调整
			.----------------------------------------------*)
			IF axHorMovingBtn_M[iAxisId] AND (NOT axHorMovingBtn_G[iAxisId]) AND (NOT xLimit_Left) THEN
				(*左*)
				alrTotalAdjust_Horz[iAxisId]:= alrTotalAdjust_Horz[iAxisId]-
				i_lrVel_HorzAdjust*	MAJOR_TSK_CYCLE_TIME*1;

				axHorMoving_G[iAxisId]:= FALSE;
				axHorMoving_M[iAxisId]:= TRUE;
			ELSIF axHorMovingBtn_G[iAxisId] AND (NOT axHorMovingBtn_M[iAxisId]) AND (NOT xLimit_Right)  THEN
				(*右*)
				alrTotalAdjust_Horz[iAxisId]:= alrTotalAdjust_Horz[iAxisId]+
				i_lrVel_HorzAdjust*	MAJOR_TSK_CYCLE_TIME*1;

				axHorMoving_M[iAxisId]:= FALSE;
				axHorMoving_G[iAxisId]:= TRUE;
			ELSE

				axHorMoving_M[iAxisId]:= FALSE;
				axHorMoving_G[iAxisId]:= FALSE;

// 			ELSIF (NOT  axHorMovingBtn_G[iAxisId])  AND
// 				(NOT axHorMovingBtn_M[iAxisId]) AND
// 				(NOT axStopManuMove_Horz[iAxisId]) THEN
// 				axStopManuMove_Horz[iAxisId]:= TRUE;
// 				axHorMoving_M[iAxisId]:= FALSE;
// 				axHorMoving_G[iAxisId]:= FALSE;
// 				alrTotalAdjust_Horz[iAxisId]:= i_alrTarp_PrfPos[iAxisId]*
// 						pstStUnitParam^.uiDen_Horz*1000.0*pstStUnitParam^.rScrewPitch_Horz/
// 						GC_LRMOTORPPR_TRAP/UINT_TO_LREAL(pstStUnitParam^.uiNum_Horz);
// 				IF pstStUnitParam^.xMotRev_Horiz_ THEN
// 					alrTotalAdjust_Horz[iAxisId]:= -alrTotalAdjust_Horz[iAxisId];
// 				END_IF
			END_IF

			(*---------------------------2017-08-14 15:21:18
			/.横向限位处理
			.----------------------------------------------*)
			IF axHorMovingLimit_M[iAxisId] THEN(*操作侧*)
				axHorMoving_M[iAxisId]:= FALSE;
			END_IF

			IF axHorMovingLimit_G[iAxisId] THEN(*传动侧*)
				axHorMoving_G[iAxisId]:= FALSE;
			END_IF

			(*急停停止横向输出|2022.5.11.171513*)
			IF i_pstStSysParam^.xFlag_EStoping OR i_pstStSysParam^.xFlag_Estop THEN
				axHorMoving_M[iAxisId]:= FALSE;
				axHorMoving_G[iAxisId]:= FALSE;
			END_IF

			(*将操作侧和传动侧信号输出*)
			(*电机输出是按照正转和反转@一般情况正反手机电机的旋转方向是一致的即,都是向操作侧或者都是向传动侧
			我们定义正传是向操作侧@反转是向传动侧*)
			pstStIOMap_Axis_FLEXO^.o_xHorzMotor_CW:=axHorMoving_M[iAxisId];
			pstStIOMap_Axis_FLEXO^.o_xHorzMotor_CCW:=axHorMoving_G[iAxisId];
			//2023.9.25.174830确定输出方向
			o_alrTotalAdjust_Horz[iAxisId]:= alrTotalAdjust_Horz[iAxisId];
			IF pstStUnitParam^.xMotRev_Horiz_ THEN
				o_alrTotalAdjust_Horz[iAxisId]:= -o_alrTotalAdjust_Horz[iAxisId];
			END_IF
		END_FOR
	ELSE;
	END_IF
ELSE
	;
END_IF

(* ---- KS_FB_GrpHorzAdjustCtrl.st ---- *)
(*@CES
Name=KS_FB_GrpHorzAdjustCtrl
Type=FunctionBlock
TypeGuid=6f9dac99-8de1-4efc-8465-68ac443b7d08
Guid=d9626d7c-8ffe-4608-b3df-e1f14e3ddbf7
HasDeclaration=True
HasImplementation=True
*)
{DECLARATION}
FUNCTION_BLOCK KS_FB_GrpHorzAdjustCtrl
(*2023.3.8.222916
将KS_FB_AxisHorAdj屏蔽移动到KS_FB_GrpHorAdj中执行*)
(*处理了常规横向控制方式的方向控制逻辑@尝试统一方向|
@所有操作用户只关心站在套印面的左右*)
(*2025.2.7.163457 横向重复值支持整机输入*)
(*2025.2.7.170536 横向报警实现代码调整位置*)
VAR_INPUT
	i_xEn									: BOOL;(*使能*)
	i_iGrpId: INT;
	i_iGrpAxisNum_Pu						: INT; (*色组轴数*)
	i_abyGrpAxisList							: ARRAY [1..MAX_UNIT_NUM] OF BYTE; (*系的轴列表*)
	i_pastStIOMap_AxisBasic					: POINTER TO ARRAY [1..MAX_UNIT_NUM] OF StIOMap_Axis_FE; (*基础io|*)
	i_pastStIOMap_AxisExtra					: POINTER TO ARRAY [1..MAX_UNIT_NUM] OF StIOMap_Axis_Extra_FE; (* 扩展io|*)
	i_pstStSysParam: POINTER TO StSysParam;
	i_xDebugTestRun							: BOOL;
	i_xDebugTestResult_Wr					: BOOL;
	i_iDebugNum								: INT;
	i_diDebugPulse							: DINT;
	i_lrDebugPulse_PosAct					: LREAL;
	i_pastStDigitalMicroStepDrive			: POINTER TO ARRAY [1..MAX_UNIT_NUM] OF StDigitalMicroStepDrive;
	i_lrVel_HorzAdjust						: LREAL;(*mm/s; um/ms; 横向调整速度|*)
	i_lrVel_HorzPreRegister					: LREAL;(*mm/s;横向预套准速度|*)
	i_pastStAxisRapidAdjProf_H				: POINTER TO ARRAY [1..MAX_UNIT_NUM] OF StAxisRapidAdjProf_H;(*纵向快速对版|*)
	i_diPreReg_RepeatVal_H					: DINT;(*横向预套准的重复值@2025.2.7.163231*)
	i_diPreReg_SetupVal_H					: DINT;(*横向预套准的重复值@2025.2.7.163231*)
	i_xHorSyncMotorCtrl: BOOL;(*横向同步电机控制*)
	i_xHorStepDriveCtrl: BOOL;(*横向采样步进电机控制*)
	i_iStepDrivePulsePRev					: INT;(*步进电机|每一圈对应的脉冲数|default.6000||*)
	i_rStepDrivePosPPulse					: REAL;(*步进电机|每个脉冲对应的位置值 mm|default.0.0002||*)
	i_xIsDebugMode:BOOL;(*调试模式*)
	i_iStepDriveSa_Vel						: INT;(*步进电机启动速度*)
	i_iStepDrivePreReg_Vel					: INT;(*z步进电机预套速度R/MIN*)
	i_iStepDriveManu_Vel					: INT;(*z步进电机手动速度R/MIN*)
	i_iStepDriveManu_Vel_Fast				: INT;(*z步进电机手动高速速度R/MIN*)
	i_iStepDriveAuto_Vel					: INT;(*步进电机自动速度R/MIN*)
	i_iStepDriveAccTime						: INT;(*步进电机加速时间*)
	i_xHor_Goal_Flag						: BOOL;(*TRUE:目标值调整标志,走到左限位以目标值+当前修正量的值;FALSE :修正量调整标志,当前修正量-前次修正量的值*)
	i_xHor_PreRegist_Flag					: BOOL;(*横向预套准标志*)
	i_xEnaTestARC_Ink:BOOL;(*空转测试使能*)
	i_xHorLimit:BOOL;(*横向限位定义修改为左右|默认是纤维定义为正反方向*)
	i_xHorManuCtrl:BOOL;(*界面横向手动修正功能*)
END_VAR
VAR_IN_OUT
	(*2025.2.7.165301+*)
	io_byBtn_HorzPreRegister_Repeat			: BYTE;(*重复值的横向按钮@界面使用|=0 不运动|=1 按照轴距离运动|=2 整机按照单个值运动*)
	io_byBtn_HorzPreRegister_Setup			: BYTE;(*目标值的横向按钮@界面使用|=0 不运动|=1 按照轴距离运动|=2 整机按照单个值运动*)
	io_abyHorzManuTrigButton: ARRAY [1..MAX_UNIT_NUM] OF BYTE; (* 横向手动按钮|转发vs可视化界面操作| *)

END_VAR
VAR_OUTPUT
	o_xEno									: BOOL;
	o_iErNo									: INT;(*0成功\-1参数失败|*)
	o_xStepDriveDebugDne					: BOOL;
	o_xHorxPreRegister_Finish				: BOOL;
	o_xHorzMotorAlarmAtLeastOne				: BOOL;(*至少一色联动轴横向报警了*)
END_VAR
VAR
	fbKS_FB_GrpHorAdj						: KS_FB_GrpHorAdj;(*传统横向电机调整*)
	fbKS_FB_Debug_Get_mmPpul				: KS_FB_Debug_Get_mmPpul;(*测量单位脉冲对应的距离功能块mm/pul*)
	lrStepDrivePosPPulse					: LREAL;
	fbKS_FB_StepDrive_H						: KS_FB_StepDrive_H;
	iN										: INT;
	iUnitId									: INT;
	//iGrp									: INT;
	aiCommAdjustMentH						: ARRAY [1..MAX_UNIT_NUM] OF INT;
	aiCommAdjustMentH_HMI					: ARRAY [1..MAX_UNIT_NUM] OF DINT;
	iRtn									: INT;(*返回的调整量值*)
	xPreFlag_Stop							: BOOL;
	diPreReg_RepeatVal_H					: DINT;(*2025.2.7.163638+*)

// 	xFlag_Stop_In:ARRAY[1..2] OF BOOL;(*停机标志*)
// 	xFlag_Estop_In:ARRAY[1..2] OF BOOL;(*急停标志*)
// 	xFlag_Print_In:ARRAY[1..2] OF BOOL;(*印刷标志*)
// 	xLinkage_In:ARRAY[1..MAX_UNIT_NUM] OF BOOL;(*联动*)
// 	xSts_HorzPreRegister_In:ARRAY[1..2] OF BOOL;(*横向预套准状态*)
// 	xMode_HorzPreRegister_In:ARRAY[1..2] OF BOOL;(*横向预套准方式|false为设定值；true为重复值*)
// 	xBtn_HorzPreRegister_Repeat_In:ARRAY[1..2] OF BOOL;(*横向重复值按钮*)
// 	xBtn_HorzPreRegister_Setup_In:ARRAY[1..2] OF BOOL;(*横向设置值按钮*)
// 	diPreReg_RepeatVal_H_In:ARRAY[1..MAX_UNIT_NUM] OF DINT;(*横向重复值-预套准*)
// 	xFlag_HorzPreRegister_All_end_In:ARRAY[1..2] OF BOOL;(*横向预套准完成*)
// 	xHorzMotor_Alarm_In:ARRAY[1..MAX_UNIT_NUM] OF BOOL;(*横向报警*)

	xFlag_Stop_In: BOOL;(*停机标志*)
	xFlag_Estop_In: BOOL;(*急停标志*)
	xFlag_Print_In: BOOL;(*印刷标志*)
	xLinkage_In:ARRAY[1..MAX_UNIT_NUM] OF BOOL;(*联动*)
	xSts_HorzPreRegister_In:  BOOL;(*横向预套准状态*)
	xMode_HorzPreRegister_In: BOOL;(*横向预套准方式|false为设定值；true为重复值*)
	xBtn_HorzPreRegister_Repeat_In: BOOL;(*横向重复值按钮*)
	xBtn_HorzPreRegister_Setup_In: BOOL;(*横向设置值按钮*)
	diPreReg_RepeatVal_H_In:ARRAY[1..MAX_UNIT_NUM] OF DINT;(*横向重复值-预套准*)
	xFlag_HorzPreRegister_All_end_In:BOOL;(*横向预套准完成*)
	xHorzMotor_Alarm_In:ARRAY[1..MAX_UNIT_NUM] OF BOOL;(*横向报警*)

END_VAR

{IMPLEMENTATION}
Action_Input();
Action_Act();
Action_Output();
